(* IEC 61131-3 sources: plc-st-coding-agent/progress/evidence/f14_v13_self_20261113/jobs/custom_deepseek-v4pro, 102 files *)

(* ---- public-easy-01.candidate_01.st ---- *)
(*
ENGINEERING_CONTRACT
Pump_Motor: activation=rising edge bottleSensor (PUB001); hold until finishedButton rising edge cycle reset (PUB008); does not stop on later step starts; BOOL latch.
Filling_Valve: activation=rising edge cleaningConfirmButton (PUB002); hold until finishedButton rising (PUB008); BOOL latch.
Capping_Machine: activation=rising edge fillingConfirmButton (PUB003); hold until finishedButton rising (PUB008); BOOL latch.
Packing_Machine: activation=rising edge cappingConfirmButton (PUB004); hold until finishedButton rising (PUB008); BOOL latch.
Completion_Light: activation=rising edge packingConfirmButton (PUB005/PUB006); hold until finishedButton rising (PUB007/PUB008); BOOL latch.
Priority: finishedButton reset overrides same-scan set edges. Inputs are edge-triggered; no interlock between buttons is specified.
*)

(* CONTRACT_RULES [
{"kind":"hold_until_reset","output":"Pump_Motor","set_input":"bottleSensor","reset_input":"finishedButton"},
{"kind":"hold_until_reset","output":"Filling_Valve","set_input":"cleaningConfirmButton","reset_input":"finishedButton"},
{"kind":"hold_until_reset","output":"Capping_Machine","set_input":"fillingConfirmButton","reset_input":"finishedButton"},
{"kind":"hold_until_reset","output":"Packing_Machine","set_input":"cappingConfirmButton","reset_input":"finishedButton"},
{"kind":"hold_until_reset","output":"Completion_Light","set_input":"packingConfirmButton","reset_input":"finishedButton"}
] *)

FUNCTION_BLOCK AutomatedFillingLineControl
VAR_INPUT
    bottleSensor : BOOL;
    cleaningConfirmButton : BOOL;
    fillingConfirmButton : BOOL;
    cappingConfirmButton : BOOL;
    packingConfirmButton : BOOL;
    finishedButton : BOOL;
END_VAR
VAR_OUTPUT
    Pump_Motor : BOOL;
    Filling_Valve : BOOL;
    Capping_Machine : BOOL;
    Packing_Machine : BOOL;
    Completion_Light : BOOL;
END_VAR
VAR
    pump_latch : BOOL := FALSE;
    fill_latch : BOOL := FALSE;
    cap_latch : BOOL := FALSE;
    pack_latch : BOOL := FALSE;
    light_latch : BOOL := FALSE;

    trigBottle : R_TRIG;
    trigClean : R_TRIG;
    trigFill : R_TRIG;
    trigCap : R_TRIG;
    trigPack : R_TRIG;
    trigFinished : R_TRIG;

    tmp_bottle_edge : BOOL;
    tmp_clean_edge : BOOL;
    tmp_fill_edge : BOOL;
    tmp_cap_edge : BOOL;
    tmp_pack_edge : BOOL;
    tmp_finished_edge : BOOL;
END_VAR

trigBottle(CLK := bottleSensor);
tmp_bottle_edge := trigBottle.Q;

trigClean(CLK := cleaningConfirmButton);
tmp_clean_edge := trigClean.Q;

trigFill(CLK := fillingConfirmButton);
tmp_fill_edge := trigFill.Q;

trigCap(CLK := cappingConfirmButton);
tmp_cap_edge := trigCap.Q;

trigPack(CLK := packingConfirmButton);
tmp_pack_edge := trigPack.Q;

trigFinished(CLK := finishedButton);
tmp_finished_edge := trigFinished.Q;

IF tmp_finished_edge THEN
    pump_latch := FALSE;
    fill_latch := FALSE;
    cap_latch := FALSE;
    pack_latch := FALSE;
    light_latch := FALSE;
ELSE
    IF tmp_bottle_edge THEN
        pump_latch := TRUE;
    END_IF;

    IF tmp_clean_edge THEN
        fill_latch := TRUE;
    END_IF;

    IF tmp_fill_edge THEN
        cap_latch := TRUE;
    END_IF;

    IF tmp_cap_edge THEN
        pack_latch := TRUE;
    END_IF;

    IF tmp_pack_edge THEN
        light_latch := TRUE;
    END_IF;
END_IF;

Pump_Motor := pump_latch;
Filling_Valve := fill_latch;
Capping_Machine := cap_latch;
Packing_Machine := pack_latch;
Completion_Light := light_latch;

END_FUNCTION_BLOCK

(* ---- public-easy-01.candidate_02.st ---- *)
(*
ENGINEERING_CONTRACT
Pump_Motor: activation=rising edge bottleSensor (PUB001); hold until finishedButton rising edge cycle reset (PUB008); does not stop on later step starts; BOOL latch.
Filling_Valve: activation=rising edge cleaningConfirmButton (PUB002); hold until finishedButton rising (PUB008); BOOL latch.
Capping_Machine: activation=rising edge fillingConfirmButton (PUB003); hold until finishedButton rising (PUB008); BOOL latch.
Packing_Machine: activation=rising edge cappingConfirmButton (PUB004); hold until finishedButton rising (PUB008); BOOL latch.
Completion_Light: activation=rising edge packingConfirmButton (PUB005/PUB006); hold until finishedButton rising (PUB007/PUB008); BOOL latch.
Priority: finishedButton reset overrides same-scan set edges. Inputs are edge-triggered; no interlock between buttons is specified.
*)

(* CONTRACT_RULES [
{"kind":"hold_until_reset","output":"Pump_Motor","set_input":"bottleSensor","reset_input":"finishedButton"},
{"kind":"hold_until_reset","output":"Filling_Valve","set_input":"cleaningConfirmButton","reset_input":"finishedButton"},
{"kind":"hold_until_reset","output":"Capping_Machine","set_input":"fillingConfirmButton","reset_input":"finishedButton"},
{"kind":"hold_until_reset","output":"Packing_Machine","set_input":"cappingConfirmButton","reset_input":"finishedButton"},
{"kind":"hold_until_reset","output":"Completion_Light","set_input":"packingConfirmButton","reset_input":"finishedButton"}
] *)

FUNCTION_BLOCK AutomatedFillingLineControl
VAR_INPUT
    bottleSensor : BOOL;
    cleaningConfirmButton : BOOL;
    fillingConfirmButton : BOOL;
    cappingConfirmButton : BOOL;
    packingConfirmButton : BOOL;
    finishedButton : BOOL;
END_VAR
VAR_OUTPUT
    Pump_Motor : BOOL;
    Filling_Valve : BOOL;
    Capping_Machine : BOOL;
    Packing_Machine : BOOL;
    Completion_Light : BOOL;
END_VAR
VAR
    pump_latch : BOOL := FALSE;
    fill_latch : BOOL := FALSE;
    cap_latch : BOOL := FALSE;
    pack_latch : BOOL := FALSE;
    light_latch : BOOL := FALSE;

    trigBottle : R_TRIG;
    trigClean : R_TRIG;
    trigFill : R_TRIG;
    trigCap : R_TRIG;
    trigPack : R_TRIG;
    trigFinished : R_TRIG;

    tmp_bottle_edge : BOOL;
    tmp_clean_edge : BOOL;
    tmp_fill_edge : BOOL;
    tmp_cap_edge : BOOL;
    tmp_pack_edge : BOOL;
    tmp_finished_edge : BOOL;
END_VAR

trigBottle(CLK := bottleSensor);
tmp_bottle_edge := trigBottle.Q;

trigClean(CLK := cleaningConfirmButton);
tmp_clean_edge := trigClean.Q;

trigFill(CLK := fillingConfirmButton);
tmp_fill_edge := trigFill.Q;

trigCap(CLK := cappingConfirmButton);
tmp_cap_edge := trigCap.Q;

trigPack(CLK := packingConfirmButton);
tmp_pack_edge := trigPack.Q;

trigFinished(CLK := finishedButton);
tmp_finished_edge := trigFinished.Q;

IF tmp_finished_edge THEN
    pump_latch := FALSE;
    fill_latch := FALSE;
    cap_latch := FALSE;
    pack_latch := FALSE;
    light_latch := FALSE;
ELSE
    IF tmp_bottle_edge THEN
        pump_latch := TRUE;
    END_IF;

    IF tmp_clean_edge AND pump_latch THEN
        fill_latch := TRUE;
    END_IF;

    IF tmp_fill_edge AND fill_latch THEN
        cap_latch := TRUE;
    END_IF;

    IF tmp_cap_edge AND cap_latch THEN
        pack_latch := TRUE;
    END_IF;

    IF tmp_pack_edge AND pack_latch THEN
        light_latch := TRUE;
    END_IF;
END_IF;

Pump_Motor := pump_latch;
Filling_Valve := fill_latch;
Capping_Machine := cap_latch;
Packing_Machine := pack_latch;
Completion_Light := light_latch;

END_FUNCTION_BLOCK

(* ---- public-easy-01.candidate_03.st ---- *)
(*
ENGINEERING_CONTRACT
Pump_Motor: activation=rising edge bottleSensor (PUB001); hold until finishedButton rising edge cycle reset (PUB008); does not stop on later step starts; BOOL latch.
Filling_Valve: activation=rising edge cleaningConfirmButton (PUB002); hold until finishedButton rising (PUB008); BOOL latch.
Capping_Machine: activation=rising edge fillingConfirmButton (PUB003); hold until finishedButton rising (PUB008); BOOL latch.
Packing_Machine: activation=rising edge cappingConfirmButton (PUB004); hold until finishedButton rising (PUB008); BOOL latch.
Completion_Light: activation=rising edge packingConfirmButton (PUB005/PUB006); hold until finishedButton rising (PUB007/PUB008); BOOL latch.
Priority: finishedButton reset overrides same-scan set edges. Inputs are edge-triggered; no interlock between buttons is specified.
*)

(* CONTRACT_RULES [] *)

FUNCTION_BLOCK AutomatedFillingLineControl
VAR_INPUT
    bottleSensor : BOOL;
    cleaningConfirmButton : BOOL;
    fillingConfirmButton : BOOL;
    cappingConfirmButton : BOOL;
    packingConfirmButton : BOOL;
    finishedButton : BOOL;
END_VAR
VAR_OUTPUT
    Pump_Motor : BOOL;
    Filling_Valve : BOOL;
    Capping_Machine : BOOL;
    Packing_Machine : BOOL;
    Completion_Light : BOOL;
END_VAR
VAR
    pump_latch : BOOL := FALSE;
    fill_latch : BOOL := FALSE;
    cap_latch : BOOL := FALSE;
    pack_latch : BOOL := FALSE;
    light_latch : BOOL := FALSE;

    trigBottle : R_TRIG;
    trigClean : R_TRIG;
    trigFill : R_TRIG;
    trigCap : R_TRIG;
    trigPack : R_TRIG;
    trigFinished : R_TRIG;

    tmp_bottle_edge : BOOL;
    tmp_clean_edge : BOOL;
    tmp_fill_edge : BOOL;
    tmp_cap_edge : BOOL;
    tmp_pack_edge : BOOL;
    tmp_finished_edge : BOOL;
END_VAR

trigBottle(CLK := bottleSensor);
tmp_bottle_edge := trigBottle.Q;

trigClean(CLK := cleaningConfirmButton);
tmp_clean_edge := trigClean.Q;

trigFill(CLK := fillingConfirmButton);
tmp_fill_edge := trigFill.Q;

trigCap(CLK := cappingConfirmButton);
tmp_cap_edge := trigCap.Q;

trigPack(CLK := packingConfirmButton);
tmp_pack_edge := trigPack.Q;

trigFinished(CLK := finishedButton);
tmp_finished_edge := trigFinished.Q;

IF tmp_finished_edge THEN
    pump_latch := FALSE;
    fill_latch := FALSE;
    cap_latch := FALSE;
    pack_latch := FALSE;
    light_latch := FALSE;
ELSE
    IF tmp_bottle_edge THEN
        pump_latch := TRUE;
    END_IF;

    IF tmp_clean_edge AND pump_latch THEN
        fill_latch := TRUE;
    END_IF;

    IF tmp_fill_edge AND fill_latch THEN
        cap_latch := TRUE;
    END_IF;

    IF tmp_cap_edge AND cap_latch THEN
        pack_latch := TRUE;
    END_IF;

    IF tmp_pack_edge AND pack_latch THEN
        light_latch := TRUE;
    END_IF;
END_IF;

Pump_Motor := pump_latch;
Filling_Valve := fill_latch;
Capping_Machine := cap_latch;
Packing_Machine := pack_latch;
Completion_Light := light_latch;

END_FUNCTION_BLOCK

(* ---- public-easy-01.candidate_04.st ---- *)
(*
ENGINEERING_CONTRACT
Pump_Motor: activation=rising edge bottleSensor (PUB001); hold until finishedButton rising edge cycle reset (PUB008); does not stop on later step starts; BOOL latch.
Filling_Valve: activation=rising edge cleaningConfirmButton (PUB002); hold until finishedButton rising (PUB008); BOOL latch.
Capping_Machine: activation=rising edge fillingConfirmButton (PUB003); hold until finishedButton rising (PUB008); BOOL latch.
Packing_Machine: activation=rising edge cappingConfirmButton (PUB004); hold until finishedButton rising (PUB008); BOOL latch.
Completion_Light: activation=rising edge packingConfirmButton (PUB005/PUB006); hold until finishedButton rising (PUB007/PUB008); BOOL latch.
Priority: finishedButton reset overrides same-scan set edges. Inputs are edge-triggered; no interlock between buttons is specified.
*)

(* CONTRACT_RULES [] *)

FUNCTION_BLOCK AutomatedFillingLineControl
VAR_INPUT
    bottleSensor : BOOL;
    cleaningConfirmButton : BOOL;
    fillingConfirmButton : BOOL;
    cappingConfirmButton : BOOL;
    packingConfirmButton : BOOL;
    finishedButton : BOOL;
END_VAR
VAR_OUTPUT
    Pump_Motor : BOOL;
    Filling_Valve : BOOL;
    Capping_Machine : BOOL;
    Packing_Machine : BOOL;
    Completion_Light : BOOL;
END_VAR
VAR
    pump_latch : BOOL := FALSE;
    fill_latch : BOOL := FALSE;
    cap_latch : BOOL := FALSE;
    pack_latch : BOOL := FALSE;
    light_latch : BOOL := FALSE;

    trigBottle : R_TRIG;
    trigClean : R_TRIG;
    trigFill : R_TRIG;
    trigCap : R_TRIG;
    trigPack : R_TRIG;
    trigFinished : R_TRIG;

    tmp_bottle_edge : BOOL;
    tmp_clean_edge : BOOL;
    tmp_fill_edge : BOOL;
    tmp_cap_edge : BOOL;
    tmp_pack_edge : BOOL;
    tmp_finished_edge : BOOL;
END_VAR

trigBottle(CLK := bottleSensor);
tmp_bottle_edge := trigBottle.Q;

trigClean(CLK := cleaningConfirmButton);
tmp_clean_edge := trigClean.Q;

trigFill(CLK := fillingConfirmButton);
tmp_fill_edge := trigFill.Q;

trigCap(CLK := cappingConfirmButton);
tmp_cap_edge := trigCap.Q;

trigPack(CLK := packingConfirmButton);
tmp_pack_edge := trigPack.Q;

trigFinished(CLK := finishedButton);
tmp_finished_edge := trigFinished.Q;

IF finishedButton THEN
    pump_latch := FALSE;
    fill_latch := FALSE;
    cap_latch := FALSE;
    pack_latch := FALSE;
    light_latch := FALSE;
ELSE
    IF tmp_bottle_edge THEN
        pump_latch := TRUE;
    END_IF;

    IF tmp_clean_edge THEN
        fill_latch := TRUE;
    END_IF;

    IF tmp_fill_edge THEN
        cap_latch := TRUE;
    END_IF;

    IF tmp_cap_edge THEN
        pack_latch := TRUE;
    END_IF;

    IF tmp_pack_edge THEN
        light_latch := TRUE;
    END_IF;
END_IF;

Pump_Motor := pump_latch;
Filling_Valve := fill_latch;
Capping_Machine := cap_latch;
Packing_Machine := pack_latch;
Completion_Light := light_latch;

END_FUNCTION_BLOCK

(* ---- public-easy-01.patch_base_02.st ---- *)
(*
ENGINEERING_CONTRACT
Pump_Motor: activation=rising edge bottleSensor (PUB001); hold until finishedButton rising edge cycle reset (PUB008); does not stop on later step starts; BOOL latch.
Filling_Valve: activation=rising edge cleaningConfirmButton (PUB002); hold until finishedButton rising (PUB008); BOOL latch.
Capping_Machine: activation=rising edge fillingConfirmButton (PUB003); hold until finishedButton rising (PUB008); BOOL latch.
Packing_Machine: activation=rising edge cappingConfirmButton (PUB004); hold until finishedButton rising (PUB008); BOOL latch.
Completion_Light: activation=rising edge packingConfirmButton (PUB005/PUB006); hold until finishedButton rising (PUB007/PUB008); BOOL latch.
Priority: finishedButton reset overrides same-scan set edges. Inputs are edge-triggered; no interlock between buttons is specified.
*)

(* CONTRACT_RULES [
{"kind":"hold_until_reset","output":"Pump_Motor","set_input":"bottleSensor","reset_input":"finishedButton"},
{"kind":"hold_until_reset","output":"Filling_Valve","set_input":"cleaningConfirmButton","reset_input":"finishedButton"},
{"kind":"hold_until_reset","output":"Capping_Machine","set_input":"fillingConfirmButton","reset_input":"finishedButton"},
{"kind":"hold_until_reset","output":"Packing_Machine","set_input":"cappingConfirmButton","reset_input":"finishedButton"},
{"kind":"hold_until_reset","output":"Completion_Light","set_input":"packingConfirmButton","reset_input":"finishedButton"}
] *)

FUNCTION_BLOCK AutomatedFillingLineControl
VAR_INPUT
    bottleSensor : BOOL;
    cleaningConfirmButton : BOOL;
    fillingConfirmButton : BOOL;
    cappingConfirmButton : BOOL;
    packingConfirmButton : BOOL;
    finishedButton : BOOL;
END_VAR
VAR_OUTPUT
    Pump_Motor : BOOL;
    Filling_Valve : BOOL;
    Capping_Machine : BOOL;
    Packing_Machine : BOOL;
    Completion_Light : BOOL;
END_VAR
VAR
    pump_latch : BOOL := FALSE;
    fill_latch : BOOL := FALSE;
    cap_latch : BOOL := FALSE;
    pack_latch : BOOL := FALSE;
    light_latch : BOOL := FALSE;

    trigBottle : R_TRIG;
    trigClean : R_TRIG;
    trigFill : R_TRIG;
    trigCap : R_TRIG;
    trigPack : R_TRIG;
    trigFinished : R_TRIG;

    tmp_bottle_edge : BOOL;
    tmp_clean_edge : BOOL;
    tmp_fill_edge : BOOL;
    tmp_cap_edge : BOOL;
    tmp_pack_edge : BOOL;
    tmp_finished_edge : BOOL;
END_VAR

trigBottle(CLK := bottleSensor);
tmp_bottle_edge := trigBottle.Q;

trigClean(CLK := cleaningConfirmButton);
tmp_clean_edge := trigClean.Q;

trigFill(CLK := fillingConfirmButton);
tmp_fill_edge := trigFill.Q;

trigCap(CLK := cappingConfirmButton);
tmp_cap_edge := trigCap.Q;

trigPack(CLK := packingConfirmButton);
tmp_pack_edge := trigPack.Q;

trigFinished(CLK := finishedButton);
tmp_finished_edge := trigFinished.Q;

IF tmp_finished_edge THEN
    pump_latch := FALSE;
    fill_latch := FALSE;
    cap_latch := FALSE;
    pack_latch := FALSE;
    light_latch := FALSE;
ELSE
    IF tmp_bottle_edge THEN
        pump_latch := TRUE;
    END_IF;

    IF tmp_clean_edge THEN
        fill_latch := TRUE;
    END_IF;

    IF tmp_fill_edge THEN
        cap_latch := TRUE;
    END_IF;

    IF tmp_cap_edge THEN
        pack_latch := TRUE;
    END_IF;

    IF tmp_pack_edge THEN
        light_latch := TRUE;
    END_IF;
END_IF;

Pump_Motor := pump_latch;
Filling_Valve := fill_latch;
Capping_Machine := cap_latch;
Packing_Machine := pack_latch;
Completion_Light := light_latch;

END_FUNCTION_BLOCK

(* ---- public-easy-01.patch_base_03.st ---- *)
(*
ENGINEERING_CONTRACT
Pump_Motor: activation=rising edge bottleSensor (PUB001); hold until finishedButton rising edge cycle reset (PUB008); does not stop on later step starts; BOOL latch.
Filling_Valve: activation=rising edge cleaningConfirmButton (PUB002); hold until finishedButton rising (PUB008); BOOL latch.
Capping_Machine: activation=rising edge fillingConfirmButton (PUB003); hold until finishedButton rising (PUB008); BOOL latch.
Packing_Machine: activation=rising edge cappingConfirmButton (PUB004); hold until finishedButton rising (PUB008); BOOL latch.
Completion_Light: activation=rising edge packingConfirmButton (PUB005/PUB006); hold until finishedButton rising (PUB007/PUB008); BOOL latch.
Priority: finishedButton reset overrides same-scan set edges. Inputs are edge-triggered; no interlock between buttons is specified.
*)

(* CONTRACT_RULES [
{"kind":"hold_until_reset","output":"Pump_Motor","set_input":"bottleSensor","reset_input":"finishedButton"},
{"kind":"hold_until_reset","output":"Filling_Valve","set_input":"cleaningConfirmButton","reset_input":"finishedButton"},
{"kind":"hold_until_reset","output":"Capping_Machine","set_input":"fillingConfirmButton","reset_input":"finishedButton"},
{"kind":"hold_until_reset","output":"Packing_Machine","set_input":"cappingConfirmButton","reset_input":"finishedButton"},
{"kind":"hold_until_reset","output":"Completion_Light","set_input":"packingConfirmButton","reset_input":"finishedButton"}
] *)

FUNCTION_BLOCK AutomatedFillingLineControl
VAR_INPUT
    bottleSensor : BOOL;
    cleaningConfirmButton : BOOL;
    fillingConfirmButton : BOOL;
    cappingConfirmButton : BOOL;
    packingConfirmButton : BOOL;
    finishedButton : BOOL;
END_VAR
VAR_OUTPUT
    Pump_Motor : BOOL;
    Filling_Valve : BOOL;
    Capping_Machine : BOOL;
    Packing_Machine : BOOL;
    Completion_Light : BOOL;
END_VAR
VAR
    pump_latch : BOOL := FALSE;
    fill_latch : BOOL := FALSE;
    cap_latch : BOOL := FALSE;
    pack_latch : BOOL := FALSE;
    light_latch : BOOL := FALSE;

    trigBottle : R_TRIG;
    trigClean : R_TRIG;
    trigFill : R_TRIG;
    trigCap : R_TRIG;
    trigPack : R_TRIG;
    trigFinished : R_TRIG;

    tmp_bottle_edge : BOOL;
    tmp_clean_edge : BOOL;
    tmp_fill_edge : BOOL;
    tmp_cap_edge : BOOL;
    tmp_pack_edge : BOOL;
    tmp_finished_edge : BOOL;
END_VAR

trigBottle(CLK := bottleSensor);
tmp_bottle_edge := trigBottle.Q;

trigClean(CLK := cleaningConfirmButton);
tmp_clean_edge := trigClean.Q;

trigFill(CLK := fillingConfirmButton);
tmp_fill_edge := trigFill.Q;

trigCap(CLK := cappingConfirmButton);
tmp_cap_edge := trigCap.Q;

trigPack(CLK := packingConfirmButton);
tmp_pack_edge := trigPack.Q;

trigFinished(CLK := finishedButton);
tmp_finished_edge := trigFinished.Q;

IF tmp_finished_edge THEN
    pump_latch := FALSE;
    fill_latch := FALSE;
    cap_latch := FALSE;
    pack_latch := FALSE;
    light_latch := FALSE;
ELSE
    IF tmp_bottle_edge THEN
        pump_latch := TRUE;
    END_IF;

    IF tmp_clean_edge AND pump_latch THEN
        fill_latch := TRUE;
    END_IF;

    IF tmp_fill_edge AND fill_latch THEN
        cap_latch := TRUE;
    END_IF;

    IF tmp_cap_edge AND cap_latch THEN
        pack_latch := TRUE;
    END_IF;

    IF tmp_pack_edge AND pack_latch THEN
        light_latch := TRUE;
    END_IF;
END_IF;

Pump_Motor := pump_latch;
Filling_Valve := fill_latch;
Capping_Machine := cap_latch;
Packing_Machine := pack_latch;
Completion_Light := light_latch;

END_FUNCTION_BLOCK

(* ---- public-easy-01.patch_base_04.st ---- *)
(*
ENGINEERING_CONTRACT
Pump_Motor: activation=rising edge bottleSensor (PUB001); hold until finishedButton rising edge cycle reset (PUB008); does not stop on later step starts; BOOL latch.
Filling_Valve: activation=rising edge cleaningConfirmButton (PUB002); hold until finishedButton rising (PUB008); BOOL latch.
Capping_Machine: activation=rising edge fillingConfirmButton (PUB003); hold until finishedButton rising (PUB008); BOOL latch.
Packing_Machine: activation=rising edge cappingConfirmButton (PUB004); hold until finishedButton rising (PUB008); BOOL latch.
Completion_Light: activation=rising edge packingConfirmButton (PUB005/PUB006); hold until finishedButton rising (PUB007/PUB008); BOOL latch.
Priority: finishedButton reset overrides same-scan set edges. Inputs are edge-triggered; no interlock between buttons is specified.
*)

(* CONTRACT_RULES [] *)

FUNCTION_BLOCK AutomatedFillingLineControl
VAR_INPUT
    bottleSensor : BOOL;
    cleaningConfirmButton : BOOL;
    fillingConfirmButton : BOOL;
    cappingConfirmButton : BOOL;
    packingConfirmButton : BOOL;
    finishedButton : BOOL;
END_VAR
VAR_OUTPUT
    Pump_Motor : BOOL;
    Filling_Valve : BOOL;
    Capping_Machine : BOOL;
    Packing_Machine : BOOL;
    Completion_Light : BOOL;
END_VAR
VAR
    pump_latch : BOOL := FALSE;
    fill_latch : BOOL := FALSE;
    cap_latch : BOOL := FALSE;
    pack_latch : BOOL := FALSE;
    light_latch : BOOL := FALSE;

    trigBottle : R_TRIG;
    trigClean : R_TRIG;
    trigFill : R_TRIG;
    trigCap : R_TRIG;
    trigPack : R_TRIG;
    trigFinished : R_TRIG;

    tmp_bottle_edge : BOOL;
    tmp_clean_edge : BOOL;
    tmp_fill_edge : BOOL;
    tmp_cap_edge : BOOL;
    tmp_pack_edge : BOOL;
    tmp_finished_edge : BOOL;
END_VAR

trigBottle(CLK := bottleSensor);
tmp_bottle_edge := trigBottle.Q;

trigClean(CLK := cleaningConfirmButton);
tmp_clean_edge := trigClean.Q;

trigFill(CLK := fillingConfirmButton);
tmp_fill_edge := trigFill.Q;

trigCap(CLK := cappingConfirmButton);
tmp_cap_edge := trigCap.Q;

trigPack(CLK := packingConfirmButton);
tmp_pack_edge := trigPack.Q;

trigFinished(CLK := finishedButton);
tmp_finished_edge := trigFinished.Q;

IF tmp_finished_edge THEN
    pump_latch := FALSE;
    fill_latch := FALSE;
    cap_latch := FALSE;
    pack_latch := FALSE;
    light_latch := FALSE;
ELSE
    IF tmp_bottle_edge THEN
        pump_latch := TRUE;
    END_IF;

    IF tmp_clean_edge AND pump_latch THEN
        fill_latch := TRUE;
    END_IF;

    IF tmp_fill_edge AND fill_latch THEN
        cap_latch := TRUE;
    END_IF;

    IF tmp_cap_edge AND cap_latch THEN
        pack_latch := TRUE;
    END_IF;

    IF tmp_pack_edge AND pack_latch THEN
        light_latch := TRUE;
    END_IF;
END_IF;

Pump_Motor := pump_latch;
Filling_Valve := fill_latch;
Capping_Machine := cap_latch;
Packing_Machine := pack_latch;
Completion_Light := light_latch;

END_FUNCTION_BLOCK

(* ---- public-easy-01.raw_candidate_01.st ---- *)
(*
ENGINEERING_CONTRACT
Pump_Motor: activation=rising edge bottleSensor (PUB001); hold until finishedButton rising edge cycle reset (PUB008); does not stop on later step starts; BOOL latch.
Filling_Valve: activation=rising edge cleaningConfirmButton (PUB002); hold until finishedButton rising (PUB008); BOOL latch.
Capping_Machine: activation=rising edge fillingConfirmButton (PUB003); hold until finishedButton rising (PUB008); BOOL latch.
Packing_Machine: activation=rising edge cappingConfirmButton (PUB004); hold until finishedButton rising (PUB008); BOOL latch.
Completion_Light: activation=rising edge packingConfirmButton (PUB005/PUB006); hold until finishedButton rising (PUB007/PUB008); BOOL latch.
Priority: finishedButton reset overrides same-scan set edges. Inputs are edge-triggered; no interlock between buttons is specified.
*)

(* CONTRACT_RULES [
{"kind":"hold_until_reset","output":"Pump_Motor","set_input":"bottleSensor","reset_input":"finishedButton"},
{"kind":"hold_until_reset","output":"Filling_Valve","set_input":"cleaningConfirmButton","reset_input":"finishedButton"},
{"kind":"hold_until_reset","output":"Capping_Machine","set_input":"fillingConfirmButton","reset_input":"finishedButton"},
{"kind":"hold_until_reset","output":"Packing_Machine","set_input":"cappingConfirmButton","reset_input":"finishedButton"},
{"kind":"hold_until_reset","output":"Completion_Light","set_input":"packingConfirmButton","reset_input":"finishedButton"}
] *)

FUNCTION_BLOCK AutomatedFillingLineControl
VAR_INPUT
    bottleSensor : BOOL;
    cleaningConfirmButton : BOOL;
    fillingConfirmButton : BOOL;
    cappingConfirmButton : BOOL;
    packingConfirmButton : BOOL;
    finishedButton : BOOL;
END_VAR
VAR_OUTPUT
    Pump_Motor : BOOL;
    Filling_Valve : BOOL;
    Capping_Machine : BOOL;
    Packing_Machine : BOOL;
    Completion_Light : BOOL;
END_VAR
VAR
    pump_latch : BOOL := FALSE;
    fill_latch : BOOL := FALSE;
    cap_latch : BOOL := FALSE;
    pack_latch : BOOL := FALSE;
    light_latch : BOOL := FALSE;

    trigBottle : R_TRIG;
    trigClean : R_TRIG;
    trigFill : R_TRIG;
    trigCap : R_TRIG;
    trigPack : R_TRIG;
    trigFinished : R_TRIG;

    tmp_bottle_edge : BOOL;
    tmp_clean_edge : BOOL;
    tmp_fill_edge : BOOL;
    tmp_cap_edge : BOOL;
    tmp_pack_edge : BOOL;
    tmp_finished_edge : BOOL;
END_VAR

trigBottle(CLK := bottleSensor);
tmp_bottle_edge := trigBottle.Q;

trigClean(CLK := cleaningConfirmButton);
tmp_clean_edge := trigClean.Q;

trigFill(CLK := fillingConfirmButton);
tmp_fill_edge := trigFill.Q;

trigCap(CLK := cappingConfirmButton);
tmp_cap_edge := trigCap.Q;

trigPack(CLK := packingConfirmButton);
tmp_pack_edge := trigPack.Q;

trigFinished(CLK := finishedButton);
tmp_finished_edge := trigFinished.Q;

IF tmp_finished_edge THEN
    pump_latch := FALSE;
    fill_latch := FALSE;
    cap_latch := FALSE;
    pack_latch := FALSE;
    light_latch := FALSE;
ELSE
    IF tmp_bottle_edge THEN
        pump_latch := TRUE;
    END_IF;

    IF tmp_clean_edge THEN
        fill_latch := TRUE;
    END_IF;

    IF tmp_fill_edge THEN
        cap_latch := TRUE;
    END_IF;

    IF tmp_cap_edge THEN
        pack_latch := TRUE;
    END_IF;

    IF tmp_pack_edge THEN
        light_latch := TRUE;
    END_IF;
END_IF;

Pump_Motor := pump_latch;
Filling_Valve := fill_latch;
Capping_Machine := cap_latch;
Packing_Machine := pack_latch;
Completion_Light := light_latch;

END_FUNCTION_BLOCK

(* ---- public-easy-01.raw_candidate_02.st ---- *)
(*
ENGINEERING_CONTRACT
Pump_Motor: activation=rising edge bottleSensor (PUB001); hold until finishedButton rising edge cycle reset (PUB008); does not stop on later step starts; BOOL latch.
Filling_Valve: activation=rising edge cleaningConfirmButton (PUB002); hold until finishedButton rising (PUB008); BOOL latch.
Capping_Machine: activation=rising edge fillingConfirmButton (PUB003); hold until finishedButton rising (PUB008); BOOL latch.
Packing_Machine: activation=rising edge cappingConfirmButton (PUB004); hold until finishedButton rising (PUB008); BOOL latch.
Completion_Light: activation=rising edge packingConfirmButton (PUB005/PUB006); hold until finishedButton rising (PUB007/PUB008); BOOL latch.
Priority: finishedButton reset overrides same-scan set edges. Inputs are edge-triggered; no interlock between buttons is specified.
*)

(* CONTRACT_RULES [
{"kind":"hold_until_reset","output":"Pump_Motor","set_input":"bottleSensor","reset_input":"finishedButton"},
{"kind":"hold_until_reset","output":"Filling_Valve","set_input":"cleaningConfirmButton","reset_input":"finishedButton"},
{"kind":"hold_until_reset","output":"Capping_Machine","set_input":"fillingConfirmButton","reset_input":"finishedButton"},
{"kind":"hold_until_reset","output":"Packing_Machine","set_input":"cappingConfirmButton","reset_input":"finishedButton"},
{"kind":"hold_until_reset","output":"Completion_Light","set_input":"packingConfirmButton","reset_input":"finishedButton"}
] *)

FUNCTION_BLOCK AutomatedFillingLineControl
VAR_INPUT
    bottleSensor : BOOL;
    cleaningConfirmButton : BOOL;
    fillingConfirmButton : BOOL;
    cappingConfirmButton : BOOL;
    packingConfirmButton : BOOL;
    finishedButton : BOOL;
END_VAR
VAR_OUTPUT
    Pump_Motor : BOOL;
    Filling_Valve : BOOL;
    Capping_Machine : BOOL;
    Packing_Machine : BOOL;
    Completion_Light : BOOL;
END_VAR
VAR
    pump_latch : BOOL := FALSE;
    fill_latch : BOOL := FALSE;
    cap_latch : BOOL := FALSE;
    pack_latch : BOOL := FALSE;
    light_latch : BOOL := FALSE;

    trigBottle : R_TRIG;
    trigClean : R_TRIG;
    trigFill : R_TRIG;
    trigCap : R_TRIG;
    trigPack : R_TRIG;
    trigFinished : R_TRIG;

    tmp_bottle_edge : BOOL;
    tmp_clean_edge : BOOL;
    tmp_fill_edge : BOOL;
    tmp_cap_edge : BOOL;
    tmp_pack_edge : BOOL;
    tmp_finished_edge : BOOL;
END_VAR

trigBottle(CLK := bottleSensor);
tmp_bottle_edge := trigBottle.Q;

trigClean(CLK := cleaningConfirmButton);
tmp_clean_edge := trigClean.Q;

trigFill(CLK := fillingConfirmButton);
tmp_fill_edge := trigFill.Q;

trigCap(CLK := cappingConfirmButton);
tmp_cap_edge := trigCap.Q;

trigPack(CLK := packingConfirmButton);
tmp_pack_edge := trigPack.Q;

trigFinished(CLK := finishedButton);
tmp_finished_edge := trigFinished.Q;

IF tmp_finished_edge THEN
    pump_latch := FALSE;
    fill_latch := FALSE;
    cap_latch := FALSE;
    pack_latch := FALSE;
    light_latch := FALSE;
ELSE
    IF tmp_bottle_edge THEN
        pump_latch := TRUE;
    END_IF;

    IF tmp_clean_edge AND pump_latch THEN
        fill_latch := TRUE;
    END_IF;

    IF tmp_fill_edge AND fill_latch THEN
        cap_latch := TRUE;
    END_IF;

    IF tmp_cap_edge AND cap_latch THEN
        pack_latch := TRUE;
    END_IF;

    IF tmp_pack_edge AND pack_latch THEN
        light_latch := TRUE;
    END_IF;
END_IF;

Pump_Motor := pump_latch;
Filling_Valve := fill_latch;
Capping_Machine := cap_latch;
Packing_Machine := pack_latch;
Completion_Light := light_latch;

END_FUNCTION_BLOCK

(* ---- public-easy-01.raw_candidate_03.st ---- *)
(*
ENGINEERING_CONTRACT
Pump_Motor: activation=rising edge bottleSensor (PUB001); hold until finishedButton rising edge cycle reset (PUB008); does not stop on later step starts; BOOL latch.
Filling_Valve: activation=rising edge cleaningConfirmButton (PUB002); hold until finishedButton rising (PUB008); BOOL latch.
Capping_Machine: activation=rising edge fillingConfirmButton (PUB003); hold until finishedButton rising (PUB008); BOOL latch.
Packing_Machine: activation=rising edge cappingConfirmButton (PUB004); hold until finishedButton rising (PUB008); BOOL latch.
Completion_Light: activation=rising edge packingConfirmButton (PUB005/PUB006); hold until finishedButton rising (PUB007/PUB008); BOOL latch.
Priority: finishedButton reset overrides same-scan set edges. Inputs are edge-triggered; no interlock between buttons is specified.
*)

(* CONTRACT_RULES [] *)

FUNCTION_BLOCK AutomatedFillingLineControl
VAR_INPUT
    bottleSensor : BOOL;
    cleaningConfirmButton : BOOL;
    fillingConfirmButton : BOOL;
    cappingConfirmButton : BOOL;
    packingConfirmButton : BOOL;
    finishedButton : BOOL;
END_VAR
VAR_OUTPUT
    Pump_Motor : BOOL;
    Filling_Valve : BOOL;
    Capping_Machine : BOOL;
    Packing_Machine : BOOL;
    Completion_Light : BOOL;
END_VAR
VAR
    pump_latch : BOOL := FALSE;
    fill_latch : BOOL := FALSE;
    cap_latch : BOOL := FALSE;
    pack_latch : BOOL := FALSE;
    light_latch : BOOL := FALSE;

    trigBottle : R_TRIG;
    trigClean : R_TRIG;
    trigFill : R_TRIG;
    trigCap : R_TRIG;
    trigPack : R_TRIG;
    trigFinished : R_TRIG;

    tmp_bottle_edge : BOOL;
    tmp_clean_edge : BOOL;
    tmp_fill_edge : BOOL;
    tmp_cap_edge : BOOL;
    tmp_pack_edge : BOOL;
    tmp_finished_edge : BOOL;
END_VAR

trigBottle(CLK := bottleSensor);
tmp_bottle_edge := trigBottle.Q;

trigClean(CLK := cleaningConfirmButton);
tmp_clean_edge := trigClean.Q;

trigFill(CLK := fillingConfirmButton);
tmp_fill_edge := trigFill.Q;

trigCap(CLK := cappingConfirmButton);
tmp_cap_edge := trigCap.Q;

trigPack(CLK := packingConfirmButton);
tmp_pack_edge := trigPack.Q;

trigFinished(CLK := finishedButton);
tmp_finished_edge := trigFinished.Q;

IF tmp_finished_edge THEN
    pump_latch := FALSE;
    fill_latch := FALSE;
    cap_latch := FALSE;
    pack_latch := FALSE;
    light_latch := FALSE;
ELSE
    IF tmp_bottle_edge THEN
        pump_latch := TRUE;
    END_IF;

    IF tmp_clean_edge AND pump_latch THEN
        fill_latch := TRUE;
    END_IF;

    IF tmp_fill_edge AND fill_latch THEN
        cap_latch := TRUE;
    END_IF;

    IF tmp_cap_edge AND cap_latch THEN
        pack_latch := TRUE;
    END_IF;

    IF tmp_pack_edge AND pack_latch THEN
        light_latch := TRUE;
    END_IF;
END_IF;

Pump_Motor := pump_latch;
Filling_Valve := fill_latch;
Capping_Machine := cap_latch;
Packing_Machine := pack_latch;
Completion_Light := light_latch;

END_FUNCTION_BLOCK

(* ---- public-easy-01.raw_candidate_04.st ---- *)
(*
ENGINEERING_CONTRACT
Pump_Motor: activation=rising edge bottleSensor (PUB001); hold until finishedButton rising edge cycle reset (PUB008); does not stop on later step starts; BOOL latch.
Filling_Valve: activation=rising edge cleaningConfirmButton (PUB002); hold until finishedButton rising (PUB008); BOOL latch.
Capping_Machine: activation=rising edge fillingConfirmButton (PUB003); hold until finishedButton rising (PUB008); BOOL latch.
Packing_Machine: activation=rising edge cappingConfirmButton (PUB004); hold until finishedButton rising (PUB008); BOOL latch.
Completion_Light: activation=rising edge packingConfirmButton (PUB005/PUB006); hold until finishedButton rising (PUB007/PUB008); BOOL latch.
Priority: finishedButton reset overrides same-scan set edges. Inputs are edge-triggered; no interlock between buttons is specified.
*)

(* CONTRACT_RULES [] *)

FUNCTION_BLOCK AutomatedFillingLineControl
VAR_INPUT
    bottleSensor : BOOL;
    cleaningConfirmButton : BOOL;
    fillingConfirmButton : BOOL;
    cappingConfirmButton : BOOL;
    packingConfirmButton : BOOL;
    finishedButton : BOOL;
END_VAR
VAR_OUTPUT
    Pump_Motor : BOOL;
    Filling_Valve : BOOL;
    Capping_Machine : BOOL;
    Packing_Machine : BOOL;
    Completion_Light : BOOL;
END_VAR
VAR
    pump_latch : BOOL := FALSE;
    fill_latch : BOOL := FALSE;
    cap_latch : BOOL := FALSE;
    pack_latch : BOOL := FALSE;
    light_latch : BOOL := FALSE;

    trigBottle : R_TRIG;
    trigClean : R_TRIG;
    trigFill : R_TRIG;
    trigCap : R_TRIG;
    trigPack : R_TRIG;
    trigFinished : R_TRIG;

    tmp_bottle_edge : BOOL;
    tmp_clean_edge : BOOL;
    tmp_fill_edge : BOOL;
    tmp_cap_edge : BOOL;
    tmp_pack_edge : BOOL;
    tmp_finished_edge : BOOL;
END_VAR

trigBottle(CLK := bottleSensor);
tmp_bottle_edge := trigBottle.Q;

trigClean(CLK := cleaningConfirmButton);
tmp_clean_edge := trigClean.Q;

trigFill(CLK := fillingConfirmButton);
tmp_fill_edge := trigFill.Q;

trigCap(CLK := cappingConfirmButton);
tmp_cap_edge := trigCap.Q;

trigPack(CLK := packingConfirmButton);
tmp_pack_edge := trigPack.Q;

trigFinished(CLK := finishedButton);
tmp_finished_edge := trigFinished.Q;

IF finishedButton THEN
    pump_latch := FALSE;
    fill_latch := FALSE;
    cap_latch := FALSE;
    pack_latch := FALSE;
    light_latch := FALSE;
ELSE
    IF tmp_bottle_edge THEN
        pump_latch := TRUE;
    END_IF;

    IF tmp_clean_edge THEN
        fill_latch := TRUE;
    END_IF;

    IF tmp_fill_edge THEN
        cap_latch := TRUE;
    END_IF;

    IF tmp_cap_edge THEN
        pack_latch := TRUE;
    END_IF;

    IF tmp_pack_edge THEN
        light_latch := TRUE;
    END_IF;
END_IF;

Pump_Motor := pump_latch;
Filling_Valve := fill_latch;
Capping_Machine := cap_latch;
Packing_Machine := pack_latch;
Completion_Light := light_latch;

END_FUNCTION_BLOCK

(* ---- public-easy-02.candidate_01.st ---- *)
(* ENGINEERING_CONTRACT
- previousValue: internal DWORD state, retains last processed value across cycles; first call establishes baseline and emits no edges.
- hasChanged: activation = value <> previousValue after first scan; no retention; automatically false next scan when equal.
- hasRisingEdges/risingBits/noOfRisingBits: activation = bits transition 0->1 from previousValue to value; no retention; counts 0..32.
- hasFallingEdges/fallingBits/noOfFallingBits: activation = bits transition 1->0; no retention; counts 0..32.
- Same-scan: rising and falling may both be true for different bit positions; hasChanged is true if either set.
- Units/boundaries: 32-bit DWORD masks, USINT counts range 0..32; detection each scan after first. PUB001.
*)
(* CONTRACT_RULES [] *)
FUNCTION_BLOCK FB
VAR_INPUT
    value : DWORD;
END_VAR
VAR_OUTPUT
    hasChanged : BOOL;
    hasRisingEdges : BOOL;
    risingBits : DWORD;
    noOfRisingBits : USINT;
    hasFallingEdges : BOOL;
    fallingBits : DWORD;
    noOfFallingBits : USINT;
END_VAR
VAR
    previousValue : DWORD;
    hasPrevious : BOOL := FALSE;
    tmp_changed : DWORD;
    tmp_rising : DWORD;
    tmp_falling : DWORD;
    tmp_i : UDINT;
    tmp_count : USINT;
END_VAR

IF NOT hasPrevious THEN
    previousValue := value;
    hasPrevious := TRUE;
    hasChanged := FALSE;
    hasRisingEdges := FALSE;
    risingBits := DWORD#0;
    noOfRisingBits := 0;
    hasFallingEdges := FALSE;
    fallingBits := DWORD#0;
    noOfFallingBits := 0;
    RETURN;
END_IF;

tmp_changed := value XOR previousValue;
tmp_rising := value AND (NOT previousValue);
tmp_falling := previousValue AND (NOT value);

hasChanged := tmp_changed <> DWORD#0;
hasRisingEdges := tmp_rising <> DWORD#0;
hasFallingEdges := tmp_falling <> DWORD#0;

risingBits := tmp_rising;
fallingBits := tmp_falling;

tmp_count := 0;
FOR tmp_i := 0 TO 31 DO
    IF (risingBits AND SHL(DWORD#1, tmp_i)) <> DWORD#0 THEN
        tmp_count := tmp_count + 1;
    END_IF;
END_FOR;
noOfRisingBits := tmp_count;

tmp_count := 0;
FOR tmp_i := 0 TO 31 DO
    IF (fallingBits AND SHL(DWORD#1, tmp_i)) <> DWORD#0 THEN
        tmp_count := tmp_count + 1;
    END_IF;
END_FOR;
noOfFallingBits := tmp_count;

previousValue := value;
END_FUNCTION_BLOCK

(* ---- public-easy-02.candidate_02.st ---- *)
(* ENGINEERING_CONTRACT
- previousValue: internal DWORD state initialized to DWORD#0; first cycle detects edges relative to 0, so every set bit is a rising edge. PUB001.
- hasChanged: activation = value <> previousValue after first scan; no retention; automatically false next scan when equal.
- hasRisingEdges/risingBits/noOfRisingBits: activation = bits transition 0->1 from previousValue to value; no retention; counts 0..32.
- hasFallingEdges/fallingBits/noOfFallingBits: activation = bits transition 1->0; no retention; counts 0..32.
- Same-scan: rising and falling may both be true for different bit positions; hasChanged is true if either set.
- Units/boundaries: 32-bit DWORD masks, USINT counts range 0..32; detection each scan after first. PUB001.
*)
(* CONTRACT_RULES [] *)
FUNCTION_BLOCK FB
VAR_INPUT
    value : DWORD;
END_VAR
VAR_OUTPUT
    hasChanged : BOOL;
    hasRisingEdges : BOOL;
    risingBits : DWORD;
    noOfRisingBits : USINT;
    hasFallingEdges : BOOL;
    fallingBits : DWORD;
    noOfFallingBits : USINT;
END_VAR
VAR
    previousValue : DWORD;
    tmp_changed : DWORD;
    tmp_rising : DWORD;
    tmp_falling : DWORD;
    tmp_i : UDINT;
    tmp_count : USINT;
END_VAR

tmp_changed := value XOR previousValue;
tmp_rising := value AND (NOT previousValue);
tmp_falling := previousValue AND (NOT value);

hasChanged := tmp_changed <> DWORD#0;
hasRisingEdges := tmp_rising <> DWORD#0;
hasFallingEdges := tmp_falling <> DWORD#0;

risingBits := tmp_rising;
fallingBits := tmp_falling;

tmp_count := 0;
FOR tmp_i := 0 TO 31 DO
    IF (risingBits AND SHL(DWORD#1, tmp_i)) <> DWORD#0 THEN
        tmp_count := tmp_count + 1;
    END_IF;
END_FOR;
noOfRisingBits := tmp_count;

tmp_count := 0;
FOR tmp_i := 0 TO 31 DO
    IF (fallingBits AND SHL(DWORD#1, tmp_i)) <> DWORD#0 THEN
        tmp_count := tmp_count + 1;
    END_IF;
END_FOR;
noOfFallingBits := tmp_count;

previousValue := value;
END_FUNCTION_BLOCK

(* ---- public-easy-02.patch_base_02.st ---- *)
(* ENGINEERING_CONTRACT
- previousValue: internal DWORD state, retains last processed value across cycles; first call establishes baseline and emits no edges.
- hasChanged: activation = value <> previousValue after first scan; no retention; automatically false next scan when equal.
- hasRisingEdges/risingBits/noOfRisingBits: activation = bits transition 0->1 from previousValue to value; no retention; counts 0..32.
- hasFallingEdges/fallingBits/noOfFallingBits: activation = bits transition 1->0; no retention; counts 0..32.
- Same-scan: rising and falling may both be true for different bit positions; hasChanged is true if either set.
- Units/boundaries: 32-bit DWORD masks, USINT counts range 0..32; detection each scan after first. PUB001.
*)
(* CONTRACT_RULES [] *)
FUNCTION_BLOCK FB
VAR_INPUT
    value : DWORD;
END_VAR
VAR_OUTPUT
    hasChanged : BOOL;
    hasRisingEdges : BOOL;
    risingBits : DWORD;
    noOfRisingBits : USINT;
    hasFallingEdges : BOOL;
    fallingBits : DWORD;
    noOfFallingBits : USINT;
END_VAR
VAR
    previousValue : DWORD;
    hasPrevious : BOOL := FALSE;
    tmp_changed : DWORD;
    tmp_rising : DWORD;
    tmp_falling : DWORD;
    tmp_i : UDINT;
    tmp_count : USINT;
END_VAR

IF NOT hasPrevious THEN
    previousValue := value;
    hasPrevious := TRUE;
    hasChanged := FALSE;
    hasRisingEdges := FALSE;
    risingBits := DWORD#0;
    noOfRisingBits := 0;
    hasFallingEdges := FALSE;
    fallingBits := DWORD#0;
    noOfFallingBits := 0;
    RETURN;
END_IF;

tmp_changed := value XOR previousValue;
tmp_rising := value AND (NOT previousValue);
tmp_falling := previousValue AND (NOT value);

hasChanged := tmp_changed <> DWORD#0;
hasRisingEdges := tmp_rising <> DWORD#0;
hasFallingEdges := tmp_falling <> DWORD#0;

risingBits := tmp_rising;
fallingBits := tmp_falling;

tmp_count := 0;
FOR tmp_i := 0 TO 31 DO
    IF (risingBits AND SHL(DWORD#1, tmp_i)) <> DWORD#0 THEN
        tmp_count := tmp_count + 1;
    END_IF;
END_FOR;
noOfRisingBits := tmp_count;

tmp_count := 0;
FOR tmp_i := 0 TO 31 DO
    IF (fallingBits AND SHL(DWORD#1, tmp_i)) <> DWORD#0 THEN
        tmp_count := tmp_count + 1;
    END_IF;
END_FOR;
noOfFallingBits := tmp_count;

previousValue := value;
END_FUNCTION_BLOCK

(* ---- public-easy-02.raw_candidate_01.st ---- *)
(* ENGINEERING_CONTRACT
- previousValue: internal DWORD state, retains last processed value across cycles; first call establishes baseline and emits no edges.
- hasChanged: activation = value <> previousValue after first scan; no retention; automatically false next scan when equal.
- hasRisingEdges/risingBits/noOfRisingBits: activation = bits transition 0->1 from previousValue to value; no retention; counts 0..32.
- hasFallingEdges/fallingBits/noOfFallingBits: activation = bits transition 1->0; no retention; counts 0..32.
- Same-scan: rising and falling may both be true for different bit positions; hasChanged is true if either set.
- Units/boundaries: 32-bit DWORD masks, USINT counts range 0..32; detection each scan after first. PUB001.
*)
(* CONTRACT_RULES [] *)
FUNCTION_BLOCK FB
VAR_INPUT
    value : DWORD;
END_VAR
VAR_OUTPUT
    hasChanged : BOOL;
    hasRisingEdges : BOOL;
    risingBits : DWORD;
    noOfRisingBits : USINT;
    hasFallingEdges : BOOL;
    fallingBits : DWORD;
    noOfFallingBits : USINT;
END_VAR
VAR
    previousValue : DWORD;
    hasPrevious : BOOL := FALSE;
    tmp_changed : DWORD;
    tmp_rising : DWORD;
    tmp_falling : DWORD;
    tmp_i : UDINT;
    tmp_count : USINT;
END_VAR

IF NOT hasPrevious THEN
    previousValue := value;
    hasPrevious := TRUE;
    hasChanged := FALSE;
    hasRisingEdges := FALSE;
    risingBits := DWORD#0;
    noOfRisingBits := 0;
    hasFallingEdges := FALSE;
    fallingBits := DWORD#0;
    noOfFallingBits := 0;
    RETURN;
END_IF;

tmp_changed := value XOR previousValue;
tmp_rising := value AND (NOT previousValue);
tmp_falling := previousValue AND (NOT value);

hasChanged := tmp_changed <> DWORD#0;
hasRisingEdges := tmp_rising <> DWORD#0;
hasFallingEdges := tmp_falling <> DWORD#0;

risingBits := tmp_rising;
fallingBits := tmp_falling;

tmp_count := 0;
FOR tmp_i := 0 TO 31 DO
    IF (risingBits AND SHL(DWORD#1, tmp_i)) <> DWORD#0 THEN
        tmp_count := tmp_count + 1;
    END_IF;
END_FOR;
noOfRisingBits := tmp_count;

tmp_count := 0;
FOR tmp_i := 0 TO 31 DO
    IF (fallingBits AND SHL(DWORD#1, tmp_i)) <> DWORD#0 THEN
        tmp_count := tmp_count + 1;
    END_IF;
END_FOR;
noOfFallingBits := tmp_count;

previousValue := value;
END_FUNCTION_BLOCK

(* ---- public-easy-02.raw_candidate_02.st ---- *)
(* ENGINEERING_CONTRACT
- previousValue: internal DWORD state initialized to DWORD#0; first cycle detects edges relative to 0, so every set bit is a rising edge. PUB001.
- hasChanged: activation = value <> previousValue after first scan; no retention; automatically false next scan when equal.
- hasRisingEdges/risingBits/noOfRisingBits: activation = bits transition 0->1 from previousValue to value; no retention; counts 0..32.
- hasFallingEdges/fallingBits/noOfFallingBits: activation = bits transition 1->0; no retention; counts 0..32.
- Same-scan: rising and falling may both be true for different bit positions; hasChanged is true if either set.
- Units/boundaries: 32-bit DWORD masks, USINT counts range 0..32; detection each scan after first. PUB001.
*)
(* CONTRACT_RULES [] *)
FUNCTION_BLOCK FB
VAR_INPUT
    value : DWORD;
END_VAR
VAR_OUTPUT
    hasChanged : BOOL;
    hasRisingEdges : BOOL;
    risingBits : DWORD;
    noOfRisingBits : USINT;
    hasFallingEdges : BOOL;
    fallingBits : DWORD;
    noOfFallingBits : USINT;
END_VAR
VAR
    previousValue : DWORD;
    tmp_changed : DWORD;
    tmp_rising : DWORD;
    tmp_falling : DWORD;
    tmp_i : UDINT;
    tmp_count : USINT;
END_VAR

tmp_changed := value XOR previousValue;
tmp_rising := value AND (NOT previousValue);
tmp_falling := previousValue AND (NOT value);

hasChanged := tmp_changed <> DWORD#0;
hasRisingEdges := tmp_rising <> DWORD#0;
hasFallingEdges := tmp_falling <> DWORD#0;

risingBits := tmp_rising;
fallingBits := tmp_falling;

tmp_count := 0;
FOR tmp_i := 0 TO 31 DO
    IF (risingBits AND SHL(DWORD#1, tmp_i)) <> DWORD#0 THEN
        tmp_count := tmp_count + 1;
    END_IF;
END_FOR;
noOfRisingBits := tmp_count;

tmp_count := 0;
FOR tmp_i := 0 TO 31 DO
    IF (fallingBits AND SHL(DWORD#1, tmp_i)) <> DWORD#0 THEN
        tmp_count := tmp_count + 1;
    END_IF;
END_FOR;
noOfFallingBits := tmp_count;

previousValue := value;
END_FUNCTION_BLOCK

(* ---- public-easy-03.candidate_01.st ---- *)
(* ENGINEERING_CONTRACT
   [PUB001-PUB004] hiAlarm/loAlarm are retained hysteresis states.
   hiAlarm activates on Value>hiLevel when off; resets only on Value<hiLevel-hystWindow when on.
   loAlarm activates on Value<loLevel when off; resets only on Value>loLevel+hystWindow when on.
   Strict comparisons are used; equality causes no state change.
   Alarm outputs are not updated during configuration error; they keep their last written values.
   On first invocation alarm states default to FALSE.
   [PUB005] If loLevel>=hiLevel then error=TRUE, status=16#8001 and RETURN. This check has priority over PUB006.
   [PUB006] Else if hystWindow>=(hiLevel-loLevel) then error=TRUE, status=16#8002 and RETURN.
   Normal scan: error=FALSE, status=0, then both hysteresis states are evaluated from current Value.
   Units: REAL thresholds/hysteresis, WORD status; no timers or pulse logic.
*)
(* CONTRACT_RULES [] *)
FUNCTION_BLOCK AlarmHandling
VAR_INPUT
    Value : REAL;
    hiLevel : REAL;
    loLevel : REAL;
    hystWindow : REAL;
END_VAR
VAR_OUTPUT
    hiAlarm : BOOL;
    loAlarm : BOOL;
    error : BOOL;
    status : WORD;
END_VAR
VAR
    local_hiAlarmState : BOOL := FALSE;
    local_loAlarmState : BOOL := FALSE;
END_VAR

IF loLevel >= hiLevel THEN
    error := TRUE;
    status := 16#8001;
    RETURN;
END_IF;

IF hystWindow >= (hiLevel - loLevel) THEN
    error := TRUE;
    status := 16#8002;
    RETURN;
END_IF;

error := FALSE;
status := 0;

IF local_hiAlarmState THEN
    IF Value < (hiLevel - hystWindow) THEN
        local_hiAlarmState := FALSE;
    END_IF;
ELSE
    IF Value > hiLevel THEN
        local_hiAlarmState := TRUE;
    END_IF;
END_IF;

hiAlarm := local_hiAlarmState;

IF local_loAlarmState THEN
    IF Value > (loLevel + hystWindow) THEN
        local_loAlarmState := FALSE;
    END_IF;
ELSE
    IF Value < loLevel THEN
        local_loAlarmState := TRUE;
    END_IF;
END_IF;

loAlarm := local_loAlarmState;

END_FUNCTION_BLOCK

(* ---- public-easy-03.raw_candidate_01.st ---- *)
(* ENGINEERING_CONTRACT
   [PUB001-PUB004] hiAlarm/loAlarm are retained hysteresis states.
   hiAlarm activates on Value>hiLevel when off; resets only on Value<hiLevel-hystWindow when on.
   loAlarm activates on Value<loLevel when off; resets only on Value>loLevel+hystWindow when on.
   Strict comparisons are used; equality causes no state change.
   Alarm outputs are not updated during configuration error; they keep their last written values.
   On first invocation alarm states default to FALSE.
   [PUB005] If loLevel>=hiLevel then error=TRUE, status=16#8001 and RETURN. This check has priority over PUB006.
   [PUB006] Else if hystWindow>=(hiLevel-loLevel) then error=TRUE, status=16#8002 and RETURN.
   Normal scan: error=FALSE, status=0, then both hysteresis states are evaluated from current Value.
   Units: REAL thresholds/hysteresis, WORD status; no timers or pulse logic.
*)
(* CONTRACT_RULES [] *)
FUNCTION_BLOCK AlarmHandling
VAR_INPUT
    Value : REAL;
    hiLevel : REAL;
    loLevel : REAL;
    hystWindow : REAL;
END_VAR
VAR_OUTPUT
    hiAlarm : BOOL;
    loAlarm : BOOL;
    error : BOOL;
    status : WORD;
END_VAR
VAR
    local_hiAlarmState : BOOL := FALSE;
    local_loAlarmState : BOOL := FALSE;
END_VAR

IF loLevel >= hiLevel THEN
    error := TRUE;
    status := 16#8001;
    RETURN;
END_IF;

IF hystWindow >= (hiLevel - loLevel) THEN
    error := TRUE;
    status := 16#8002;
    RETURN;
END_IF;

error := FALSE;
status := 0;

IF local_hiAlarmState THEN
    IF Value < (hiLevel - hystWindow) THEN
        local_hiAlarmState := FALSE;
    END_IF;
ELSE
    IF Value > hiLevel THEN
        local_hiAlarmState := TRUE;
    END_IF;
END_IF;

hiAlarm := local_hiAlarmState;

IF local_loAlarmState THEN
    IF Value > (loLevel + hystWindow) THEN
        local_loAlarmState := FALSE;
    END_IF;
ELSE
    IF Value < loLevel THEN
        local_loAlarmState := TRUE;
    END_IF;
END_IF;

loAlarm := local_loAlarmState;

END_FUNCTION_BLOCK

(* ---- public-easy-04.candidate_01.st ---- *)
FUNCTION_BLOCK JamPump
(*
ENGINEERING_CONTRACT
- VFD_RUN: active only when PASTE_E_STOP_NC AND debounce valid (PUB002); off immediately on estop false or viscosity false; no retention.
- Debounce: valid only after VISCOSITY_OK continuously true for DebounceTime; input false clears valid immediately. Incomplete timing is cleared while estop false; already-valid condition is not cleared by estop.
- Runtime: PUMP_RUNTIME_ACC adds CycleTime only when final same-scan VFD_RUN is true; retained while stopped; zero at init (PUB003/PUB005).
- Maintenance: PUMP_MAINT_DUE latches when accumulated LTIME >= 500h; no reset; informational and does not influence VFD_RUN (PUB004).
- Same-scan: reset/invalidate first, compute VFD_RUN, then add runtime using final VFD_RUN.
- Units: TIME inputs converted to LTIME; comparison >=; 500h = LTIME#500h.
*)
(* CONTRACT_RULES [] *)
VAR_INPUT
    VISCOSITY_OK : BOOL;
    PASTE_E_STOP_NC : BOOL;
    DebounceTime : TIME;
    CycleTime : TIME;
END_VAR
VAR_OUTPUT
    VFD_RUN : BOOL;
    PUMP_MAINT_DUE : BOOL;
    PUMP_RUNTIME_ACC : LTIME;
END_VAR
VAR
    tmp_debounce_elapsed : LTIME := LTIME#0s;
    tmp_debounce_valid : BOOL := FALSE;
    tmp_runtime_acc : LTIME := LTIME#0s;
    tmp_maintenance_latched : BOOL := FALSE;
    tmp_cycle_lt : LTIME;
    tmp_debounce_pt_lt : LTIME;
    tmp_maint_threshold_lt : LTIME := LTIME#500h;
END_VAR

tmp_cycle_lt := TIME_TO_LTIME(CycleTime);
tmp_debounce_pt_lt := TIME_TO_LTIME(DebounceTime);

IF NOT VISCOSITY_OK THEN
    tmp_debounce_elapsed := LTIME#0s;
    tmp_debounce_valid := FALSE;
ELSIF NOT PASTE_E_STOP_NC THEN
    IF NOT tmp_debounce_valid THEN
        tmp_debounce_elapsed := LTIME#0s;
    END_IF;
ELSE
    IF NOT tmp_debounce_valid THEN
        tmp_debounce_elapsed := tmp_debounce_elapsed + tmp_cycle_lt;
        IF tmp_debounce_elapsed >= tmp_debounce_pt_lt THEN
            tmp_debounce_valid := TRUE;
            tmp_debounce_elapsed := tmp_debounce_pt_lt;
        END_IF;
    END_IF;
END_IF;

VFD_RUN := PASTE_E_STOP_NC AND tmp_debounce_valid;

IF VFD_RUN THEN
    tmp_runtime_acc := tmp_runtime_acc + tmp_cycle_lt;
END_IF;

IF tmp_runtime_acc >= tmp_maint_threshold_lt THEN
    tmp_maintenance_latched := TRUE;
END_IF;

PUMP_MAINT_DUE := tmp_maintenance_latched;
PUMP_RUNTIME_ACC := tmp_runtime_acc;

END_FUNCTION_BLOCK

(* ---- public-easy-04.candidate_02.st ---- *)
FUNCTION_BLOCK JamPump
(*
ENGINEERING_CONTRACT
- VFD_RUN: active only when PASTE_E_STOP_NC AND debounce valid (PUB002); off immediately on estop false or viscosity false; no retention.
- Debounce: valid only after VISCOSITY_OK continuously true for DebounceTime; input false clears valid immediately. Incomplete timing is cleared while estop false; already-valid condition is not cleared by estop.
- Runtime: PUMP_RUNTIME_ACC adds CycleTime only when final same-scan VFD_RUN is true; retained while stopped; zero at init (PUB003/PUB005).
- Maintenance: PUMP_MAINT_DUE latches when accumulated LTIME >= 500h; no reset; informational and does not influence VFD_RUN (PUB004).
- Same-scan: reset/invalidate first, compute VFD_RUN, then add runtime using final VFD_RUN.
- Units: TIME inputs converted to LTIME; comparison >=; 500h = LTIME#500h.
*)
(* CONTRACT_RULES [] *)
VAR_INPUT
    VISCOSITY_OK : BOOL;
    PASTE_E_STOP_NC : BOOL;
    DebounceTime : TIME;
    CycleTime : TIME;
END_VAR
VAR_OUTPUT
    VFD_RUN : BOOL;
    PUMP_MAINT_DUE : BOOL;
    PUMP_RUNTIME_ACC : LTIME;
END_VAR
VAR
    tmp_debounce_elapsed : LTIME := LTIME#0s;
    tmp_debounce_valid : BOOL := FALSE;
    tmp_runtime_acc : LTIME := LTIME#0s;
    tmp_maintenance_latched : BOOL := FALSE;
    tmp_cycle_lt : LTIME;
    tmp_debounce_pt_lt : LTIME;
    tmp_maint_threshold_lt : LTIME := LTIME#500h;
END_VAR

tmp_cycle_lt := TIME_TO_LTIME(CycleTime);
tmp_debounce_pt_lt := TIME_TO_LTIME(DebounceTime);

IF NOT VISCOSITY_OK THEN
    tmp_debounce_elapsed := LTIME#0s;
    tmp_debounce_valid := FALSE;
ELSIF NOT PASTE_E_STOP_NC THEN
    IF NOT tmp_debounce_valid THEN
        tmp_debounce_elapsed := LTIME#0s;
    END_IF;
ELSE
    IF NOT tmp_debounce_valid THEN
        tmp_debounce_elapsed := tmp_debounce_elapsed + tmp_cycle_lt;
        IF tmp_debounce_elapsed > tmp_debounce_pt_lt THEN
            tmp_debounce_valid := TRUE;
            tmp_debounce_elapsed := tmp_debounce_pt_lt;
        END_IF;
    END_IF;
END_IF;

VFD_RUN := PASTE_E_STOP_NC AND tmp_debounce_valid;

IF VFD_RUN THEN
    tmp_runtime_acc := tmp_runtime_acc + tmp_cycle_lt;
END_IF;

IF tmp_runtime_acc >= tmp_maint_threshold_lt THEN
    tmp_maintenance_latched := TRUE;
END_IF;

PUMP_MAINT_DUE := tmp_maintenance_latched;
PUMP_RUNTIME_ACC := tmp_runtime_acc;

END_FUNCTION_BLOCK

(* ---- public-easy-04.patch_base_02.st ---- *)
FUNCTION_BLOCK JamPump
(*
ENGINEERING_CONTRACT
- VFD_RUN: active only when PASTE_E_STOP_NC AND debounce valid (PUB002); off immediately on estop false or viscosity false; no retention.
- Debounce: valid only after VISCOSITY_OK continuously true for DebounceTime; input false clears valid immediately. Incomplete timing is cleared while estop false; already-valid condition is not cleared by estop.
- Runtime: PUMP_RUNTIME_ACC adds CycleTime only when final same-scan VFD_RUN is true; retained while stopped; zero at init (PUB003/PUB005).
- Maintenance: PUMP_MAINT_DUE latches when accumulated LTIME >= 500h; no reset; informational and does not influence VFD_RUN (PUB004).
- Same-scan: reset/invalidate first, compute VFD_RUN, then add runtime using final VFD_RUN.
- Units: TIME inputs converted to LTIME; comparison >=; 500h = LTIME#500h.
*)
(* CONTRACT_RULES [] *)
VAR_INPUT
    VISCOSITY_OK : BOOL;
    PASTE_E_STOP_NC : BOOL;
    DebounceTime : TIME;
    CycleTime : TIME;
END_VAR
VAR_OUTPUT
    VFD_RUN : BOOL;
    PUMP_MAINT_DUE : BOOL;
    PUMP_RUNTIME_ACC : LTIME;
END_VAR
VAR
    tmp_debounce_elapsed : LTIME := LTIME#0s;
    tmp_debounce_valid : BOOL := FALSE;
    tmp_runtime_acc : LTIME := LTIME#0s;
    tmp_maintenance_latched : BOOL := FALSE;
    tmp_cycle_lt : LTIME;
    tmp_debounce_pt_lt : LTIME;
    tmp_maint_threshold_lt : LTIME := LTIME#500h;
END_VAR

tmp_cycle_lt := TIME_TO_LTIME(CycleTime);
tmp_debounce_pt_lt := TIME_TO_LTIME(DebounceTime);

IF NOT VISCOSITY_OK THEN
    tmp_debounce_elapsed := LTIME#0s;
    tmp_debounce_valid := FALSE;
ELSIF NOT PASTE_E_STOP_NC THEN
    IF NOT tmp_debounce_valid THEN
        tmp_debounce_elapsed := LTIME#0s;
    END_IF;
ELSE
    IF NOT tmp_debounce_valid THEN
        tmp_debounce_elapsed := tmp_debounce_elapsed + tmp_cycle_lt;
        IF tmp_debounce_elapsed >= tmp_debounce_pt_lt THEN
            tmp_debounce_valid := TRUE;
            tmp_debounce_elapsed := tmp_debounce_pt_lt;
        END_IF;
    END_IF;
END_IF;

VFD_RUN := PASTE_E_STOP_NC AND tmp_debounce_valid;

IF VFD_RUN THEN
    tmp_runtime_acc := tmp_runtime_acc + tmp_cycle_lt;
END_IF;

IF tmp_runtime_acc >= tmp_maint_threshold_lt THEN
    tmp_maintenance_latched := TRUE;
END_IF;

PUMP_MAINT_DUE := tmp_maintenance_latched;
PUMP_RUNTIME_ACC := tmp_runtime_acc;

END_FUNCTION_BLOCK

(* ---- public-easy-04.raw_candidate_01.st ---- *)
FUNCTION_BLOCK JamPump
(*
ENGINEERING_CONTRACT
- VFD_RUN: active only when PASTE_E_STOP_NC AND debounce valid (PUB002); off immediately on estop false or viscosity false; no retention.
- Debounce: valid only after VISCOSITY_OK continuously true for DebounceTime; input false clears valid immediately. Incomplete timing is cleared while estop false; already-valid condition is not cleared by estop.
- Runtime: PUMP_RUNTIME_ACC adds CycleTime only when final same-scan VFD_RUN is true; retained while stopped; zero at init (PUB003/PUB005).
- Maintenance: PUMP_MAINT_DUE latches when accumulated LTIME >= 500h; no reset; informational and does not influence VFD_RUN (PUB004).
- Same-scan: reset/invalidate first, compute VFD_RUN, then add runtime using final VFD_RUN.
- Units: TIME inputs converted to LTIME; comparison >=; 500h = LTIME#500h.
*)
(* CONTRACT_RULES [] *)
VAR_INPUT
    VISCOSITY_OK : BOOL;
    PASTE_E_STOP_NC : BOOL;
    DebounceTime : TIME;
    CycleTime : TIME;
END_VAR
VAR_OUTPUT
    VFD_RUN : BOOL;
    PUMP_MAINT_DUE : BOOL;
    PUMP_RUNTIME_ACC : LTIME;
END_VAR
VAR
    tmp_debounce_elapsed : LTIME := LTIME#0s;
    tmp_debounce_valid : BOOL := FALSE;
    tmp_runtime_acc : LTIME := LTIME#0s;
    tmp_maintenance_latched : BOOL := FALSE;
    tmp_cycle_lt : LTIME;
    tmp_debounce_pt_lt : LTIME;
    tmp_maint_threshold_lt : LTIME := LTIME#500h;
END_VAR

tmp_cycle_lt := TIME_TO_LTIME(CycleTime);
tmp_debounce_pt_lt := TIME_TO_LTIME(DebounceTime);

IF NOT VISCOSITY_OK THEN
    tmp_debounce_elapsed := LTIME#0s;
    tmp_debounce_valid := FALSE;
ELSIF NOT PASTE_E_STOP_NC THEN
    IF NOT tmp_debounce_valid THEN
        tmp_debounce_elapsed := LTIME#0s;
    END_IF;
ELSE
    IF NOT tmp_debounce_valid THEN
        tmp_debounce_elapsed := tmp_debounce_elapsed + tmp_cycle_lt;
        IF tmp_debounce_elapsed >= tmp_debounce_pt_lt THEN
            tmp_debounce_valid := TRUE;
            tmp_debounce_elapsed := tmp_debounce_pt_lt;
        END_IF;
    END_IF;
END_IF;

VFD_RUN := PASTE_E_STOP_NC AND tmp_debounce_valid;

IF VFD_RUN THEN
    tmp_runtime_acc := tmp_runtime_acc + tmp_cycle_lt;
END_IF;

IF tmp_runtime_acc >= tmp_maint_threshold_lt THEN
    tmp_maintenance_latched := TRUE;
END_IF;

PUMP_MAINT_DUE := tmp_maintenance_latched;
PUMP_RUNTIME_ACC := tmp_runtime_acc;

END_FUNCTION_BLOCK

(* ---- public-easy-04.raw_candidate_02.st ---- *)
FUNCTION_BLOCK JamPump
(*
ENGINEERING_CONTRACT
- VFD_RUN: active only when PASTE_E_STOP_NC AND debounce valid (PUB002); off immediately on estop false or viscosity false; no retention.
- Debounce: valid only after VISCOSITY_OK continuously true for DebounceTime; input false clears valid immediately. Incomplete timing is cleared while estop false; already-valid condition is not cleared by estop.
- Runtime: PUMP_RUNTIME_ACC adds CycleTime only when final same-scan VFD_RUN is true; retained while stopped; zero at init (PUB003/PUB005).
- Maintenance: PUMP_MAINT_DUE latches when accumulated LTIME >= 500h; no reset; informational and does not influence VFD_RUN (PUB004).
- Same-scan: reset/invalidate first, compute VFD_RUN, then add runtime using final VFD_RUN.
- Units: TIME inputs converted to LTIME; comparison >=; 500h = LTIME#500h.
*)
(* CONTRACT_RULES [] *)
VAR_INPUT
    VISCOSITY_OK : BOOL;
    PASTE_E_STOP_NC : BOOL;
    DebounceTime : TIME;
    CycleTime : TIME;
END_VAR
VAR_OUTPUT
    VFD_RUN : BOOL;
    PUMP_MAINT_DUE : BOOL;
    PUMP_RUNTIME_ACC : LTIME;
END_VAR
VAR
    tmp_debounce_elapsed : LTIME := LTIME#0s;
    tmp_debounce_valid : BOOL := FALSE;
    tmp_runtime_acc : LTIME := LTIME#0s;
    tmp_maintenance_latched : BOOL := FALSE;
    tmp_cycle_lt : LTIME;
    tmp_debounce_pt_lt : LTIME;
    tmp_maint_threshold_lt : LTIME := LTIME#500h;
END_VAR

tmp_cycle_lt := TIME_TO_LTIME(CycleTime);
tmp_debounce_pt_lt := TIME_TO_LTIME(DebounceTime);

IF NOT VISCOSITY_OK THEN
    tmp_debounce_elapsed := LTIME#0s;
    tmp_debounce_valid := FALSE;
ELSIF NOT PASTE_E_STOP_NC THEN
    IF NOT tmp_debounce_valid THEN
        tmp_debounce_elapsed := LTIME#0s;
    END_IF;
ELSE
    IF NOT tmp_debounce_valid THEN
        tmp_debounce_elapsed := tmp_debounce_elapsed + tmp_cycle_lt;
        IF tmp_debounce_elapsed > tmp_debounce_pt_lt THEN
            tmp_debounce_valid := TRUE;
            tmp_debounce_elapsed := tmp_debounce_pt_lt;
        END_IF;
    END_IF;
END_IF;

VFD_RUN := PASTE_E_STOP_NC AND tmp_debounce_valid;

IF VFD_RUN THEN
    tmp_runtime_acc := tmp_runtime_acc + tmp_cycle_lt;
END_IF;

IF tmp_runtime_acc >= tmp_maint_threshold_lt THEN
    tmp_maintenance_latched := TRUE;
END_IF;

PUMP_MAINT_DUE := tmp_maintenance_latched;
PUMP_RUNTIME_ACC := tmp_runtime_acc;

END_FUNCTION_BLOCK

(* ---- public-easy-05.candidate_01.st ---- *)
FUNCTION_BLOCK WeldGapAlarmControl
(* ENGINEERING_CONTRACT
Operator_Alert: combinational; active when Gap_Exceeded has been TRUE continuously for DebounceTime after init and no E-stop. No latch, not retained; deasserts when DeboundTimer.Q false or EStop active. PUB003/PUB004.
Weld_Soft_Start_Active: active while init timer NOT Q and EStop inactive. Deactivates on first scan where 5s init timer Q true. EStop masks; no latch. PUB002/PUB004/PUB005.
Init timer: TON always enabled from power-up; wall-clock 5s. EStop masks SoftStart but does not reset/pause init timer (unspecified).
Debounce timer: IN = Gap_Exceeded AND init done AND NOT EStopActive; resets on gap false, init, EStop. PT = DebounceTime (TIME ms). PUB002/PUB003/PUB004.
Same-scan priority: EStopActive computed first; init Q then debounce Q used same scan. Boundary: SoftStart off at first scan with InitTimer.Q true. PUB002/PUB003.
*)
VAR_INPUT
    Gap_Exceeded : BOOL;
    Weld_E_Stop_NC : BOOL;
    DebounceTime : TIME;
END_VAR
VAR_OUTPUT
    Operator_Alert : BOOL;
    Weld_Soft_Start_Active : BOOL;
END_VAR
VAR
    InitTimer : TON;
    DebounceTimer : TON;
    tmp_EStopActive : BOOL;
    tmp_InitDone : BOOL;
    tmp_DebounceEnable : BOOL;
END_VAR

(* CONTRACT_RULES [] *)

tmp_EStopActive := NOT Weld_E_Stop_NC;

InitTimer(IN := TRUE, PT := T#5S);
tmp_InitDone := InitTimer.Q;

tmp_DebounceEnable := Gap_Exceeded AND tmp_InitDone AND NOT tmp_EStopActive;
DebounceTimer(IN := tmp_DebounceEnable, PT := DebounceTime);

Operator_Alert := DebounceTimer.Q AND NOT tmp_EStopActive;
Weld_Soft_Start_Active := (NOT InitTimer.Q) AND (NOT tmp_EStopActive);

END_FUNCTION_BLOCK

(* ---- public-easy-05.raw_candidate_01.st ---- *)
FUNCTION_BLOCK WeldGapAlarmControl
(* ENGINEERING_CONTRACT
Operator_Alert: combinational; active when Gap_Exceeded has been TRUE continuously for DebounceTime after init and no E-stop. No latch, not retained; deasserts when DeboundTimer.Q false or EStop active. PUB003/PUB004.
Weld_Soft_Start_Active: active while init timer NOT Q and EStop inactive. Deactivates on first scan where 5s init timer Q true. EStop masks; no latch. PUB002/PUB004/PUB005.
Init timer: TON always enabled from power-up; wall-clock 5s. EStop masks SoftStart but does not reset/pause init timer (unspecified).
Debounce timer: IN = Gap_Exceeded AND init done AND NOT EStopActive; resets on gap false, init, EStop. PT = DebounceTime (TIME ms). PUB002/PUB003/PUB004.
Same-scan priority: EStopActive computed first; init Q then debounce Q used same scan. Boundary: SoftStart off at first scan with InitTimer.Q true. PUB002/PUB003.
*)
VAR_INPUT
    Gap_Exceeded : BOOL;
    Weld_E_Stop_NC : BOOL;
    DebounceTime : TIME;
END_VAR
VAR_OUTPUT
    Operator_Alert : BOOL;
    Weld_Soft_Start_Active : BOOL;
END_VAR
VAR
    InitTimer : TON;
    DebounceTimer : TON;
    tmp_EStopActive : BOOL;
    tmp_InitDone : BOOL;
    tmp_DebounceEnable : BOOL;
END_VAR

(* CONTRACT_RULES [] *)

tmp_EStopActive := NOT Weld_E_Stop_NC;

InitTimer(IN := TRUE, PT := T#5S);
tmp_InitDone := InitTimer.Q;

tmp_DebounceEnable := Gap_Exceeded AND tmp_InitDone AND NOT tmp_EStopActive;
DebounceTimer(IN := tmp_DebounceEnable, PT := DebounceTime);

Operator_Alert := DebounceTimer.Q AND NOT tmp_EStopActive;
Weld_Soft_Start_Active := (NOT InitTimer.Q) AND (NOT tmp_EStopActive);

END_FUNCTION_BLOCK

(* ---- public-easy-06.candidate_01.st ---- *)
FUNCTION_BLOCK AerationBlowerDelayedStart
VAR_INPUT
    DO_LOW : BOOL;
    AERATION_E_STOP_NC : BOOL;
END_VAR
VAR_OUTPUT
    BLOWER_RUN : BOOL;
    AERATION_BLOWER_CYCLE_COUNT : UINT;
END_VAR
VAR
    startTimer : TON;
    blowerRising : R_TRIG;
    tmp_initDone : BOOL := FALSE;
END_VAR

(* ENGINEERING_CONTRACT
   BLOWER_RUN: combinational enable derived from TON.Q. Activate when DO_LOW AND AERATION_E_STOP_NC
   remain TRUE for 5 s (PUB001). Deactivate immediately when either input becomes FALSE; TON IN false resets
   the timer in the same scan (PUB002). No latch or hold_until_reset.
   AERATION_BLOWER_CYCLE_COUNT: retained UINT output, initialized to 0 on first scan (PUB004).
   Increment exactly once on each FALSE->TRUE edge of BLOWER_RUN (PUB003). Unit: starts; range 0..65535.
   First-scan initialization forces BLOWER_RUN FALSE and count 0 (PUB004). No speed ramp (PUB004).
*)

(* CONTRACT_RULES [] *)

IF NOT tmp_initDone THEN
    BLOWER_RUN := FALSE;
    AERATION_BLOWER_CYCLE_COUNT := 0;
    tmp_initDone := TRUE;
END_IF;

startTimer(IN := DO_LOW AND AERATION_E_STOP_NC, PT := T#5S);
BLOWER_RUN := startTimer.Q;

blowerRising(CLK := BLOWER_RUN);
IF blowerRising.Q THEN
    AERATION_BLOWER_CYCLE_COUNT := AERATION_BLOWER_CYCLE_COUNT + 1;
END_IF;

END_FUNCTION_BLOCK

(* ---- public-easy-06.raw_candidate_01.st ---- *)
FUNCTION_BLOCK AerationBlowerDelayedStart
VAR_INPUT
    DO_LOW : BOOL;
    AERATION_E_STOP_NC : BOOL;
END_VAR
VAR_OUTPUT
    BLOWER_RUN : BOOL;
    AERATION_BLOWER_CYCLE_COUNT : UINT;
END_VAR
VAR
    startTimer : TON;
    blowerRising : R_TRIG;
    tmp_initDone : BOOL := FALSE;
END_VAR

(* ENGINEERING_CONTRACT
   BLOWER_RUN: combinational enable derived from TON.Q. Activate when DO_LOW AND AERATION_E_STOP_NC
   remain TRUE for 5 s (PUB001). Deactivate immediately when either input becomes FALSE; TON IN false resets
   the timer in the same scan (PUB002). No latch or hold_until_reset.
   AERATION_BLOWER_CYCLE_COUNT: retained UINT output, initialized to 0 on first scan (PUB004).
   Increment exactly once on each FALSE->TRUE edge of BLOWER_RUN (PUB003). Unit: starts; range 0..65535.
   First-scan initialization forces BLOWER_RUN FALSE and count 0 (PUB004). No speed ramp (PUB004).
*)

(* CONTRACT_RULES [] *)

IF NOT tmp_initDone THEN
    BLOWER_RUN := FALSE;
    AERATION_BLOWER_CYCLE_COUNT := 0;
    tmp_initDone := TRUE;
END_IF;

startTimer(IN := DO_LOW AND AERATION_E_STOP_NC, PT := T#5S);
BLOWER_RUN := startTimer.Q;

blowerRising(CLK := BLOWER_RUN);
IF blowerRising.Q THEN
    AERATION_BLOWER_CYCLE_COUNT := AERATION_BLOWER_CYCLE_COUNT + 1;
END_IF;

END_FUNCTION_BLOCK

(* ---- public-hard-01.candidate_01.st ---- *)
(*
ENGINEERING_CONTRACT
Outputs/state group | activation | retention/hold | reset/deactivation | same-scan priority | units/bounds
estop: highest priority; active-low; all outputs false and internal states/latches reset (PUB001, PUB003).
Manual valve/motor: rising button toggles local latch; held between scans; reset by estop or mode change (PUB002, PUB004-PUB005).
AutoState: idle all off; fillA A on until level>=50; fillB B on until level>=80; processMode false->mix, true->fillC C on until level>=100; mix motor on until complete signal false->true while motor running; deliver D on and retained until autoStart/estop/mode change (PUB006-PUB015).
AutoStart rising restarts at fillA and suppresses threshold transition for first scan; transitions update state before output mapping this scan.
levelSensor INT cm; thresholds use >=.
mix completion uses armed condition requiring mixMotorComplete FALSE before TRUE while in mix state.
*)
(* CONTRACT_RULES [] *)
FUNCTION_BLOCK MaterialProportioningControl
VAR CONSTANT
    AUTO_IDLE : INT := 0;
    AUTO_FILL_A : INT := 1;
    AUTO_FILL_B : INT := 2;
    AUTO_FILL_C : INT := 3;
    AUTO_MIX : INT := 4;
    AUTO_DELIVER : INT := 5;
END_VAR
VAR
    autoStartRtr : R_TRIG;
    valveAStartRtr : R_TRIG;
    valveBStartRtr : R_TRIG;
    valveCStartRtr : R_TRIG;
    valveDStartRtr : R_TRIG;
    mixMotorStartRtr : R_TRIG;

    local_prevOpeMode : BOOL := FALSE;
    local_init : BOOL := FALSE;

    local_manualA : BOOL := FALSE;
    local_manualB : BOOL := FALSE;
    local_manualC : BOOL := FALSE;
    local_manualD : BOOL := FALSE;
    local_manualMix : BOOL := FALSE;

    local_autoState : INT := AUTO_IDLE;
    local_firstAutoScan : BOOL := FALSE;
    local_mixArmed : BOOL := FALSE;

    local_autoStartEdge : BOOL;
    local_edgeA : BOOL;
    local_edgeB : BOOL;
    local_edgeC : BOOL;
    local_edgeD : BOOL;
    local_edgeMix : BOOL;
END_VAR

autoStartRtr(CLK := autoStart);
valveAStartRtr(CLK := valveAStart);
valveBStartRtr(CLK := valveBStart);
valveCStartRtr(CLK := valveCStart);
valveDStartRtr(CLK := valveDStart);
mixMotorStartRtr(CLK := mixMotorStart);

local_autoStartEdge := autoStartRtr.Q AND opeMode AND estop;
local_edgeA := valveAStartRtr.Q AND NOT opeMode AND estop;
local_edgeB := valveBStartRtr.Q AND NOT opeMode AND estop;
local_edgeC := valveCStartRtr.Q AND NOT opeMode AND estop;
local_edgeD := valveDStartRtr.Q AND NOT opeMode AND estop;
local_edgeMix := mixMotorStartRtr.Q AND NOT opeMode AND estop;

IF NOT local_init THEN
    local_prevOpeMode := opeMode;
    local_init := TRUE;
ELSIF local_prevOpeMode <> opeMode THEN
    local_prevOpeMode := opeMode;
    local_manualA := FALSE;
    local_manualB := FALSE;
    local_manualC := FALSE;
    local_manualD := FALSE;
    local_manualMix := FALSE;
    local_autoState := AUTO_IDLE;
    local_firstAutoScan := FALSE;
    local_mixArmed := FALSE;
END_IF;

IF NOT estop THEN
    valveARun := FALSE;
    valveBRun := FALSE;
    valveCRun := FALSE;
    valveDRun := FALSE;
    mixMotorRun := FALSE;

    local_manualA := FALSE;
    local_manualB := FALSE;
    local_manualC := FALSE;
    local_manualD := FALSE;
    local_manualMix := FALSE;
    local_autoState := AUTO_IDLE;
    local_firstAutoScan := FALSE;
    local_mixArmed := FALSE;
    RETURN;
END_IF;

IF opeMode THEN
    IF local_autoStartEdge THEN
        local_autoState := AUTO_FILL_A;
        local_firstAutoScan := TRUE;
        local_mixArmed := FALSE;
    END_IF;

    IF NOT local_firstAutoScan THEN
        IF local_autoState = AUTO_FILL_A THEN
            IF levelSensor >= 50 THEN
                local_autoState := AUTO_FILL_B;
            END_IF;
        ELSIF local_autoState = AUTO_FILL_B THEN
            IF levelSensor >= 80 THEN
                IF processMode THEN
                    local_autoState := AUTO_FILL_C;
                ELSE
                    local_autoState := AUTO_MIX;
                END_IF;
            END_IF;
        ELSIF local_autoState = AUTO_FILL_C THEN
            IF levelSensor >= 100 THEN
                local_autoState := AUTO_MIX;
            END_IF;
        ELSIF local_autoState = AUTO_MIX THEN
            IF local_mixArmed AND mixMotorComplete THEN
                local_autoState := AUTO_DELIVER;
            END_IF;
        END_IF;
    END_IF;

    IF local_autoState = AUTO_MIX THEN
        IF NOT mixMotorComplete THEN
            local_mixArmed := TRUE;
        END_IF;
    ELSE
        local_mixArmed := FALSE;
    END_IF;

    CASE local_autoState OF
        AUTO_IDLE:
            valveARun := FALSE;
            valveBRun := FALSE;
            valveCRun := FALSE;
            valveDRun := FALSE;
            mixMotorRun := FALSE;

        AUTO_FILL_A:
            valveARun := TRUE;
            valveBRun := FALSE;
            valveCRun := FALSE;
            valveDRun := FALSE;
            mixMotorRun := FALSE;

        AUTO_FILL_B:
            valveARun := FALSE;
            valveBRun := TRUE;
            valveCRun := FALSE;
            valveDRun := FALSE;
            mixMotorRun := FALSE;

        AUTO_FILL_C:
            valveARun := FALSE;
            valveBRun := FALSE;
            valveCRun := TRUE;
            valveDRun := FALSE;
            mixMotorRun := FALSE;

        AUTO_MIX:
            valveARun := FALSE;
            valveBRun := FALSE;
            valveCRun := FALSE;
            valveDRun := FALSE;
            mixMotorRun := TRUE;

        AUTO_DELIVER:
            valveARun := FALSE;
            valveBRun := FALSE;
            valveCRun := FALSE;
            valveDRun := TRUE;
            mixMotorRun := FALSE;
    END_CASE;

    local_firstAutoScan := FALSE;
ELSE
    IF local_edgeA THEN
        local_manualA := NOT local_manualA;
    END_IF;

    IF local_edgeB THEN
        local_manualB := NOT local_manualB;
    END_IF;

    IF local_edgeC THEN
        local_manualC := NOT local_manualC;
    END_IF;

    IF local_edgeD THEN
        local_manualD := NOT local_manualD;
    END_IF;

    IF local_edgeMix THEN
        local_manualMix := NOT local_manualMix;
    END_IF;

    valveARun := local_manualA;
    valveBRun := local_manualB;
    valveCRun := local_manualC;
    valveDRun := local_manualD;
    mixMotorRun := local_manualMix;
END_IF;
END_FUNCTION_BLOCK

(* ---- public-hard-01.candidate_02.st ---- *)
(*
ENGINEERING_CONTRACT
Outputs/state group | activation | retention/hold | reset/deactivation | same-scan priority | units/bounds
estop: highest priority; active-low; all outputs false and internal states/latches reset (PUB001, PUB003).
Manual valve/motor: rising button toggles local latch; held between scans; reset by estop or mode change (PUB002, PUB004-PUB005).
AutoState: idle all off; fillA A on until level>=50; fillB B on until level>=80; processMode false->mix, true->fillC C on until level>=100; mix motor on until complete signal false->true while motor running; deliver D on and retained until autoStart/estop/mode change (PUB006-PUB015).
AutoStart rising restarts at fillA and suppresses threshold transition for first scan; transitions update state before output mapping this scan.
levelSensor INT cm; thresholds use >=.
mix completion uses armed condition requiring mixMotorComplete FALSE before TRUE while in mix state.
*)
(* CONTRACT_RULES [] *)
FUNCTION_BLOCK MaterialProportioningControl
VAR_INPUT
    estop : BOOL;
    opeMode : BOOL;
    valveAStart : BOOL;
    valveBStart : BOOL;
    valveCStart : BOOL;
    valveDStart : BOOL;
    mixMotorStart : BOOL;
    autoStart : BOOL;
    processMode : BOOL;
    levelSensor : INT;
    mixMotorComplete : BOOL;
END_VAR
VAR_OUTPUT
    valveARun : BOOL;
    valveBRun : BOOL;
    valveCRun : BOOL;
    valveDRun : BOOL;
    mixMotorRun : BOOL;
END_VAR
VAR CONSTANT
    AUTO_IDLE : INT := 0;
    AUTO_FILL_A : INT := 1;
    AUTO_FILL_B : INT := 2;
    AUTO_FILL_C : INT := 3;
    AUTO_MIX : INT := 4;
    AUTO_DELIVER : INT := 5;
END_VAR
VAR
    autoStartRtr : R_TRIG;
    valveAStartRtr : R_TRIG;
    valveBStartRtr : R_TRIG;
    valveCStartRtr : R_TRIG;
    valveDStartRtr : R_TRIG;
    mixMotorStartRtr : R_TRIG;

    local_prevOpeMode : BOOL := FALSE;
    local_init : BOOL := FALSE;

    local_manualA : BOOL := FALSE;
    local_manualB : BOOL := FALSE;
    local_manualC : BOOL := FALSE;
    local_manualD : BOOL := FALSE;
    local_manualMix : BOOL := FALSE;

    local_autoState : INT := AUTO_IDLE;
    local_firstAutoScan : BOOL := FALSE;
    local_mixArmed : BOOL := FALSE;

    local_autoStartEdge : BOOL;
    local_edgeA : BOOL;
    local_edgeB : BOOL;
    local_edgeC : BOOL;
    local_edgeD : BOOL;
    local_edgeMix : BOOL;
END_VAR

autoStartRtr(CLK := autoStart);
valveAStartRtr(CLK := valveAStart);
valveBStartRtr(CLK := valveBStart);
valveCStartRtr(CLK := valveCStart);
valveDStartRtr(CLK := valveDStart);
mixMotorStartRtr(CLK := mixMotorStart);

local_autoStartEdge := autoStartRtr.Q AND opeMode AND estop;
local_edgeA := valveAStartRtr.Q AND NOT opeMode AND estop;
local_edgeB := valveBStartRtr.Q AND NOT opeMode AND estop;
local_edgeC := valveCStartRtr.Q AND NOT opeMode AND estop;
local_edgeD := valveDStartRtr.Q AND NOT opeMode AND estop;
local_edgeMix := mixMotorStartRtr.Q AND NOT opeMode AND estop;

IF NOT local_init THEN
    local_prevOpeMode := opeMode;
    local_init := TRUE;
ELSIF local_prevOpeMode <> opeMode THEN
    local_prevOpeMode := opeMode;
    local_manualA := FALSE;
    local_manualB := FALSE;
    local_manualC := FALSE;
    local_manualD := FALSE;
    local_manualMix := FALSE;
    local_autoState := AUTO_IDLE;
    local_firstAutoScan := FALSE;
    local_mixArmed := FALSE;
END_IF;

IF NOT estop THEN
    valveARun := FALSE;
    valveBRun := FALSE;
    valveCRun := FALSE;
    valveDRun := FALSE;
    mixMotorRun := FALSE;

    local_manualA := FALSE;
    local_manualB := FALSE;
    local_manualC := FALSE;
    local_manualD := FALSE;
    local_manualMix := FALSE;
    local_autoState := AUTO_IDLE;
    local_firstAutoScan := FALSE;
    local_mixArmed := FALSE;
    RETURN;
END_IF;

IF opeMode THEN
    IF local_autoStartEdge THEN
        local_autoState := AUTO_FILL_A;
        local_firstAutoScan := TRUE;
        local_mixArmed := FALSE;
    END_IF;

    IF NOT local_firstAutoScan THEN
        IF local_autoState = AUTO_FILL_A THEN
            IF levelSensor >= 50 THEN
                local_autoState := AUTO_FILL_B;
            END_IF;
        ELSIF local_autoState = AUTO_FILL_B THEN
            IF levelSensor >= 80 THEN
                IF processMode THEN
                    local_autoState := AUTO_FILL_C;
                ELSE
                    local_autoState := AUTO_MIX;
                END_IF;
            END_IF;
        ELSIF local_autoState = AUTO_FILL_C THEN
            IF levelSensor >= 100 THEN
                local_autoState := AUTO_MIX;
            END_IF;
        ELSIF local_autoState = AUTO_MIX THEN
            IF local_mixArmed AND mixMotorComplete THEN
                local_autoState := AUTO_DELIVER;
            END_IF;
        END_IF;
    END_IF;

    IF local_autoState = AUTO_MIX THEN
        IF NOT mixMotorComplete THEN
            local_mixArmed := TRUE;
        END_IF;
    ELSE
        local_mixArmed := FALSE;
    END_IF;

    CASE local_autoState OF
        AUTO_IDLE:
            valveARun := FALSE;
            valveBRun := FALSE;
            valveCRun := FALSE;
            valveDRun := FALSE;
            mixMotorRun := FALSE;

        AUTO_FILL_A:
            valveARun := TRUE;
            valveBRun := FALSE;
            valveCRun := FALSE;
            valveDRun := FALSE;
            mixMotorRun := FALSE;

        AUTO_FILL_B:
            valveARun := FALSE;
            valveBRun := TRUE;
            valveCRun := FALSE;
            valveDRun := FALSE;
            mixMotorRun := FALSE;

        AUTO_FILL_C:
            valveARun := FALSE;
            valveBRun := FALSE;
            valveCRun := TRUE;
            valveDRun := FALSE;
            mixMotorRun := FALSE;

        AUTO_MIX:
            valveARun := FALSE;
            valveBRun := FALSE;
            valveCRun := FALSE;
            valveDRun := FALSE;
            mixMotorRun := TRUE;

        AUTO_DELIVER:
            valveARun := FALSE;
            valveBRun := FALSE;
            valveCRun := FALSE;
            valveDRun := TRUE;
            mixMotorRun := FALSE;
    END_CASE;

    local_firstAutoScan := FALSE;
ELSE
    IF local_edgeA THEN
        local_manualA := NOT local_manualA;
    END_IF;

    IF local_edgeB THEN
        local_manualB := NOT local_manualB;
    END_IF;

    IF local_edgeC THEN
        local_manualC := NOT local_manualC;
    END_IF;

    IF local_edgeD THEN
        local_manualD := NOT local_manualD;
    END_IF;

    IF local_edgeMix THEN
        local_manualMix := NOT local_manualMix;
    END_IF;

    valveARun := local_manualA;
    valveBRun := local_manualB;
    valveCRun := local_manualC;
    valveDRun := local_manualD;
    mixMotorRun := local_manualMix;
END_IF;
END_FUNCTION_BLOCK

(* ---- public-hard-01.patch_base_02.st ---- *)
(*
ENGINEERING_CONTRACT
Outputs/state group | activation | retention/hold | reset/deactivation | same-scan priority | units/bounds
estop: highest priority; active-low; all outputs false and internal states/latches reset (PUB001, PUB003).
Manual valve/motor: rising button toggles local latch; held between scans; reset by estop or mode change (PUB002, PUB004-PUB005).
AutoState: idle all off; fillA A on until level>=50; fillB B on until level>=80; processMode false->mix, true->fillC C on until level>=100; mix motor on until complete signal false->true while motor running; deliver D on and retained until autoStart/estop/mode change (PUB006-PUB015).
AutoStart rising restarts at fillA and suppresses threshold transition for first scan; transitions update state before output mapping this scan.
levelSensor INT cm; thresholds use >=.
mix completion uses armed condition requiring mixMotorComplete FALSE before TRUE while in mix state.
*)
(* CONTRACT_RULES [] *)
FUNCTION_BLOCK MaterialProportioningControl
VAR CONSTANT
    AUTO_IDLE : INT := 0;
    AUTO_FILL_A : INT := 1;
    AUTO_FILL_B : INT := 2;
    AUTO_FILL_C : INT := 3;
    AUTO_MIX : INT := 4;
    AUTO_DELIVER : INT := 5;
END_VAR
VAR
    autoStartRtr : R_TRIG;
    valveAStartRtr : R_TRIG;
    valveBStartRtr : R_TRIG;
    valveCStartRtr : R_TRIG;
    valveDStartRtr : R_TRIG;
    mixMotorStartRtr : R_TRIG;

    local_prevOpeMode : BOOL := FALSE;
    local_init : BOOL := FALSE;

    local_manualA : BOOL := FALSE;
    local_manualB : BOOL := FALSE;
    local_manualC : BOOL := FALSE;
    local_manualD : BOOL := FALSE;
    local_manualMix : BOOL := FALSE;

    local_autoState : INT := AUTO_IDLE;
    local_firstAutoScan : BOOL := FALSE;
    local_mixArmed : BOOL := FALSE;

    local_autoStartEdge : BOOL;
    local_edgeA : BOOL;
    local_edgeB : BOOL;
    local_edgeC : BOOL;
    local_edgeD : BOOL;
    local_edgeMix : BOOL;
END_VAR

autoStartRtr(CLK := autoStart);
valveAStartRtr(CLK := valveAStart);
valveBStartRtr(CLK := valveBStart);
valveCStartRtr(CLK := valveCStart);
valveDStartRtr(CLK := valveDStart);
mixMotorStartRtr(CLK := mixMotorStart);

local_autoStartEdge := autoStartRtr.Q AND opeMode AND estop;
local_edgeA := valveAStartRtr.Q AND NOT opeMode AND estop;
local_edgeB := valveBStartRtr.Q AND NOT opeMode AND estop;
local_edgeC := valveCStartRtr.Q AND NOT opeMode AND estop;
local_edgeD := valveDStartRtr.Q AND NOT opeMode AND estop;
local_edgeMix := mixMotorStartRtr.Q AND NOT opeMode AND estop;

IF NOT local_init THEN
    local_prevOpeMode := opeMode;
    local_init := TRUE;
ELSIF local_prevOpeMode <> opeMode THEN
    local_prevOpeMode := opeMode;
    local_manualA := FALSE;
    local_manualB := FALSE;
    local_manualC := FALSE;
    local_manualD := FALSE;
    local_manualMix := FALSE;
    local_autoState := AUTO_IDLE;
    local_firstAutoScan := FALSE;
    local_mixArmed := FALSE;
END_IF;

IF NOT estop THEN
    valveARun := FALSE;
    valveBRun := FALSE;
    valveCRun := FALSE;
    valveDRun := FALSE;
    mixMotorRun := FALSE;

    local_manualA := FALSE;
    local_manualB := FALSE;
    local_manualC := FALSE;
    local_manualD := FALSE;
    local_manualMix := FALSE;
    local_autoState := AUTO_IDLE;
    local_firstAutoScan := FALSE;
    local_mixArmed := FALSE;
    RETURN;
END_IF;

IF opeMode THEN
    IF local_autoStartEdge THEN
        local_autoState := AUTO_FILL_A;
        local_firstAutoScan := TRUE;
        local_mixArmed := FALSE;
    END_IF;

    IF NOT local_firstAutoScan THEN
        IF local_autoState = AUTO_FILL_A THEN
            IF levelSensor >= 50 THEN
                local_autoState := AUTO_FILL_B;
            END_IF;
        ELSIF local_autoState = AUTO_FILL_B THEN
            IF levelSensor >= 80 THEN
                IF processMode THEN
                    local_autoState := AUTO_FILL_C;
                ELSE
                    local_autoState := AUTO_MIX;
                END_IF;
            END_IF;
        ELSIF local_autoState = AUTO_FILL_C THEN
            IF levelSensor >= 100 THEN
                local_autoState := AUTO_MIX;
            END_IF;
        ELSIF local_autoState = AUTO_MIX THEN
            IF local_mixArmed AND mixMotorComplete THEN
                local_autoState := AUTO_DELIVER;
            END_IF;
        END_IF;
    END_IF;

    IF local_autoState = AUTO_MIX THEN
        IF NOT mixMotorComplete THEN
            local_mixArmed := TRUE;
        END_IF;
    ELSE
        local_mixArmed := FALSE;
    END_IF;

    CASE local_autoState OF
        AUTO_IDLE:
            valveARun := FALSE;
            valveBRun := FALSE;
            valveCRun := FALSE;
            valveDRun := FALSE;
            mixMotorRun := FALSE;

        AUTO_FILL_A:
            valveARun := TRUE;
            valveBRun := FALSE;
            valveCRun := FALSE;
            valveDRun := FALSE;
            mixMotorRun := FALSE;

        AUTO_FILL_B:
            valveARun := FALSE;
            valveBRun := TRUE;
            valveCRun := FALSE;
            valveDRun := FALSE;
            mixMotorRun := FALSE;

        AUTO_FILL_C:
            valveARun := FALSE;
            valveBRun := FALSE;
            valveCRun := TRUE;
            valveDRun := FALSE;
            mixMotorRun := FALSE;

        AUTO_MIX:
            valveARun := FALSE;
            valveBRun := FALSE;
            valveCRun := FALSE;
            valveDRun := FALSE;
            mixMotorRun := TRUE;

        AUTO_DELIVER:
            valveARun := FALSE;
            valveBRun := FALSE;
            valveCRun := FALSE;
            valveDRun := TRUE;
            mixMotorRun := FALSE;
    END_CASE;

    local_firstAutoScan := FALSE;
ELSE
    IF local_edgeA THEN
        local_manualA := NOT local_manualA;
    END_IF;

    IF local_edgeB THEN
        local_manualB := NOT local_manualB;
    END_IF;

    IF local_edgeC THEN
        local_manualC := NOT local_manualC;
    END_IF;

    IF local_edgeD THEN
        local_manualD := NOT local_manualD;
    END_IF;

    IF local_edgeMix THEN
        local_manualMix := NOT local_manualMix;
    END_IF;

    valveARun := local_manualA;
    valveBRun := local_manualB;
    valveCRun := local_manualC;
    valveDRun := local_manualD;
    mixMotorRun := local_manualMix;
END_IF;
END_FUNCTION_BLOCK

(* ---- public-hard-01.raw_candidate_01.st ---- *)
(*
ENGINEERING_CONTRACT
Outputs/state group | activation | retention/hold | reset/deactivation | same-scan priority | units/bounds
estop: highest priority; active-low; all outputs false and internal states/latches reset (PUB001, PUB003).
Manual valve/motor: rising button toggles local latch; held between scans; reset by estop or mode change (PUB002, PUB004-PUB005).
AutoState: idle all off; fillA A on until level>=50; fillB B on until level>=80; processMode false->mix, true->fillC C on until level>=100; mix motor on until complete signal false->true while motor running; deliver D on and retained until autoStart/estop/mode change (PUB006-PUB015).
AutoStart rising restarts at fillA and suppresses threshold transition for first scan; transitions update state before output mapping this scan.
levelSensor INT cm; thresholds use >=.
mix completion uses armed condition requiring mixMotorComplete FALSE before TRUE while in mix state.
*)
(* CONTRACT_RULES [] *)
FUNCTION_BLOCK MaterialProportioningControl
VAR CONSTANT
    AUTO_IDLE : INT := 0;
    AUTO_FILL_A : INT := 1;
    AUTO_FILL_B : INT := 2;
    AUTO_FILL_C : INT := 3;
    AUTO_MIX : INT := 4;
    AUTO_DELIVER : INT := 5;
END_VAR
VAR
    autoStartRtr : R_TRIG;
    valveAStartRtr : R_TRIG;
    valveBStartRtr : R_TRIG;
    valveCStartRtr : R_TRIG;
    valveDStartRtr : R_TRIG;
    mixMotorStartRtr : R_TRIG;

    local_prevOpeMode : BOOL := FALSE;
    local_init : BOOL := FALSE;

    local_manualA : BOOL := FALSE;
    local_manualB : BOOL := FALSE;
    local_manualC : BOOL := FALSE;
    local_manualD : BOOL := FALSE;
    local_manualMix : BOOL := FALSE;

    local_autoState : INT := AUTO_IDLE;
    local_firstAutoScan : BOOL := FALSE;
    local_mixArmed : BOOL := FALSE;

    local_autoStartEdge : BOOL;
    local_edgeA : BOOL;
    local_edgeB : BOOL;
    local_edgeC : BOOL;
    local_edgeD : BOOL;
    local_edgeMix : BOOL;
END_VAR

autoStartRtr(CLK := autoStart);
valveAStartRtr(CLK := valveAStart);
valveBStartRtr(CLK := valveBStart);
valveCStartRtr(CLK := valveCStart);
valveDStartRtr(CLK := valveDStart);
mixMotorStartRtr(CLK := mixMotorStart);

local_autoStartEdge := autoStartRtr.Q AND opeMode AND estop;
local_edgeA := valveAStartRtr.Q AND NOT opeMode AND estop;
local_edgeB := valveBStartRtr.Q AND NOT opeMode AND estop;
local_edgeC := valveCStartRtr.Q AND NOT opeMode AND estop;
local_edgeD := valveDStartRtr.Q AND NOT opeMode AND estop;
local_edgeMix := mixMotorStartRtr.Q AND NOT opeMode AND estop;

IF NOT local_init THEN
    local_prevOpeMode := opeMode;
    local_init := TRUE;
ELSIF local_prevOpeMode <> opeMode THEN
    local_prevOpeMode := opeMode;
    local_manualA := FALSE;
    local_manualB := FALSE;
    local_manualC := FALSE;
    local_manualD := FALSE;
    local_manualMix := FALSE;
    local_autoState := AUTO_IDLE;
    local_firstAutoScan := FALSE;
    local_mixArmed := FALSE;
END_IF;

IF NOT estop THEN
    valveARun := FALSE;
    valveBRun := FALSE;
    valveCRun := FALSE;
    valveDRun := FALSE;
    mixMotorRun := FALSE;

    local_manualA := FALSE;
    local_manualB := FALSE;
    local_manualC := FALSE;
    local_manualD := FALSE;
    local_manualMix := FALSE;
    local_autoState := AUTO_IDLE;
    local_firstAutoScan := FALSE;
    local_mixArmed := FALSE;
    RETURN;
END_IF;

IF opeMode THEN
    IF local_autoStartEdge THEN
        local_autoState := AUTO_FILL_A;
        local_firstAutoScan := TRUE;
        local_mixArmed := FALSE;
    END_IF;

    IF NOT local_firstAutoScan THEN
        IF local_autoState = AUTO_FILL_A THEN
            IF levelSensor >= 50 THEN
                local_autoState := AUTO_FILL_B;
            END_IF;
        ELSIF local_autoState = AUTO_FILL_B THEN
            IF levelSensor >= 80 THEN
                IF processMode THEN
                    local_autoState := AUTO_FILL_C;
                ELSE
                    local_autoState := AUTO_MIX;
                END_IF;
            END_IF;
        ELSIF local_autoState = AUTO_FILL_C THEN
            IF levelSensor >= 100 THEN
                local_autoState := AUTO_MIX;
            END_IF;
        ELSIF local_autoState = AUTO_MIX THEN
            IF local_mixArmed AND mixMotorComplete THEN
                local_autoState := AUTO_DELIVER;
            END_IF;
        END_IF;
    END_IF;

    IF local_autoState = AUTO_MIX THEN
        IF NOT mixMotorComplete THEN
            local_mixArmed := TRUE;
        END_IF;
    ELSE
        local_mixArmed := FALSE;
    END_IF;

    CASE local_autoState OF
        AUTO_IDLE:
            valveARun := FALSE;
            valveBRun := FALSE;
            valveCRun := FALSE;
            valveDRun := FALSE;
            mixMotorRun := FALSE;

        AUTO_FILL_A:
            valveARun := TRUE;
            valveBRun := FALSE;
            valveCRun := FALSE;
            valveDRun := FALSE;
            mixMotorRun := FALSE;

        AUTO_FILL_B:
            valveARun := FALSE;
            valveBRun := TRUE;
            valveCRun := FALSE;
            valveDRun := FALSE;
            mixMotorRun := FALSE;

        AUTO_FILL_C:
            valveARun := FALSE;
            valveBRun := FALSE;
            valveCRun := TRUE;
            valveDRun := FALSE;
            mixMotorRun := FALSE;

        AUTO_MIX:
            valveARun := FALSE;
            valveBRun := FALSE;
            valveCRun := FALSE;
            valveDRun := FALSE;
            mixMotorRun := TRUE;

        AUTO_DELIVER:
            valveARun := FALSE;
            valveBRun := FALSE;
            valveCRun := FALSE;
            valveDRun := TRUE;
            mixMotorRun := FALSE;
    END_CASE;

    local_firstAutoScan := FALSE;
ELSE
    IF local_edgeA THEN
        local_manualA := NOT local_manualA;
    END_IF;

    IF local_edgeB THEN
        local_manualB := NOT local_manualB;
    END_IF;

    IF local_edgeC THEN
        local_manualC := NOT local_manualC;
    END_IF;

    IF local_edgeD THEN
        local_manualD := NOT local_manualD;
    END_IF;

    IF local_edgeMix THEN
        local_manualMix := NOT local_manualMix;
    END_IF;

    valveARun := local_manualA;
    valveBRun := local_manualB;
    valveCRun := local_manualC;
    valveDRun := local_manualD;
    mixMotorRun := local_manualMix;
END_IF;
END_FUNCTION_BLOCK
